(* IEC 61131-3 sources: deprecated-refusr-repo/GP/Main/samples (part 22) *)

(* ---- RND-EXPR_mouse-rusts-agues.st ---- *)
(*
This code implements a randomly grown symbolic expression:

((((!(!(!(xor(xor(IN40 | (xor(xor(IN19, IN3), IN23)), xor(xor(IN26 & IN29, !(IN6)), IN3 & IN48)), xor(xor(IN48 | IN38, !(IN41)), IN9 & IN1)))))) & true) | (xor(xor(!(IN21 & (IN50 | (IN33 & (!(!(IN10)))))), !(IN33)), IN31))) | (!(xor(xor((xor(xor(!(IN26 & (!(!(IN15)))), xor(xor((IN23 | (xor(xor(IN10, IN17), IN38))) | ((IN9 | IN7) | (IN42 & IN18)), (!(IN3)) | (!(IN26 & IN36))), xor(xor(!(IN23), (xor(xor(IN46, IN32), IN13)) | (!(IN45))), IN31))), !(xor(xor(!(xor(xor(IN29, IN29), IN17)), (IN32 | IN36) | (xor(xor(IN34, IN37), true))), xor(xor(IN48 & IN9, xor(xor(IN43, IN49), IN14)), IN2))))) | (!(((xor(xor(!(IN32), xor(xor(IN27, IN24), IN34)), IN7)) & true) | IN46)), !(IN23)), xor(xor(xor(xor((xor(xor((xor(xor(IN42, IN37), IN30)) | IN36, !(IN36)), IN31)) | (!(IN26 | (IN2 | IN28))), (!(IN14)) & (xor(xor((IN45 & IN11) | (xor(xor(IN8, IN48), IN36)), (!(IN36)) & (IN20 & IN4)), !(IN9 & IN11)))), (IN50 | (!(xor(xor(IN12, IN4), IN6)))) | (IN22 & ((IN46 & IN5) & (!(IN41))))), xor(xor(IN41, !(((IN26 & IN16) | (!(IN32))) | ((xor(xor(IN22, IN34), IN14)) & (xor(xor(IN18, IN31), IN36))))), xor(xor((IN8 | (IN9 & IN25)) & (xor(xor(!(IN41), !(IN45)), IN30 & IN43)), (!(IN18 | IN43)) | ((IN39 | IN36) & IN3)), xor(xor(IN44, (xor(xor(IN5, IN21), IN30)) | (xor(xor(IN43, IN17), IN49))), IN30)))), (!(xor(xor(IN44 & (!(IN21)), IN27), (xor(xor(IN34, IN5), IN26)) | (IN38 & IN23)))) | ((!((IN15 | IN19) | (!(IN41)))) & IN20)))))) & (((!((xor(xor(((IN40 & (!(IN13))) | ((!(IN22)) | IN28)) | (xor(xor((IN20 | IN38) & (!(IN15)), !(!(IN14))), true)), (xor(xor(xor(xor(IN5, IN3), IN26 | IN3), xor(xor(true | IN14, !(IN17)), xor(xor(IN17, IN36), IN47))), (xor(xor(IN3, IN48), IN41)) | (IN2 & IN4))) & IN40), ((!(IN6 & IN11)) & (IN26 & (IN27 | IN31))) | (IN49 & (!(xor(xor(IN27, IN28), IN2)))))) | ((xor(xor(!((IN41 | IN16) | (IN35 & IN24)), IN38), xor(xor(!(IN15 & IN10), (IN7 | IN17) | (IN38 & IN35)), xor(xor(IN41 & IN32, IN3 | IN1), !(IN20))))) & (xor(xor((xor(xor(IN6, IN30 | IN35), xor(xor(IN20, IN9), IN29))) & ((IN14 & IN14) & (IN34 | IN49)), IN15), xor(xor(true, !(IN41 & IN2)), (!(IN13)) | (IN24 | true))))))) | IN32) & (xor(xor(IN26, ((((xor(xor(xor(xor(xor(xor(IN9, IN24), IN27), IN45 | IN12), IN10 | IN19), IN7 | (IN12 & IN13)), (!(IN20)) & (!(IN2)))) | (xor(xor((IN20 | IN22) & (IN42 | false), !(IN43 & IN7)), xor(xor(!(IN49), xor(xor(IN31, IN26), IN38)), xor(xor(IN23, IN1), IN3))))) & (((!(IN4 & IN31)) | IN41) & (((xor(xor(IN34, IN47), IN25)) & (xor(xor(IN13, IN11), IN1))) & IN26))) & (!(xor(xor(xor(xor(IN50 & (IN10 | IN31), xor(xor(IN33, xor(xor(IN36, IN43), IN43)), xor(xor(IN21, IN20), IN23))), IN6), ((!(IN48)) | (IN35 & IN49)) & (xor(xor(xor(xor(IN1, IN38), IN48), !(IN17)), IN8 | IN26))), xor(xor((IN23 | IN47) | (xor(xor(IN19, IN38), IN1)), !(IN48)), xor(xor(false, xor(xor(IN31, IN1), IN6)), !(IN34))))))) & (xor(xor(IN9, xor(xor((!((IN29 & IN46) & (!(IN5)))) | IN47, (!((IN45 & IN35) & (!(IN14)))) & IN1), IN14 | (!(IN38)))), xor(xor((!(!(!(IN40)))) & ((xor(xor(!(IN18), IN7), IN17 & IN6)) | (xor(xor(xor(xor(IN12, IN34), IN21), true | IN23), !(IN1)))), !(IN43)), (((IN6 & IN32) | (!(IN11))) & (!(IN24))) & (!(xor(xor(IN36 | IN16, !(IN7)), !(IN30)))))))), (xor(xor(xor(xor((xor(xor(!(IN40 & IN14), xor(xor(!(IN45), xor(xor(IN10, IN14), IN43)), !(IN16))), xor(xor(IN10 | IN17, xor(xor(true, IN13), IN11)), IN4 & IN1))) | IN23, IN43), xor(xor(IN7, !(xor(xor(!(IN30), IN16 | IN10), IN26 | IN18))), !(!(IN42 | IN8)))), ((!(IN46)) & (xor(xor(IN45, xor(xor(!(IN32), xor(xor(IN41, IN14), IN50)), IN22 & IN33)), IN23 & IN27))) & IN4), IN2)) | (!((xor(xor(xor(xor(IN7, xor(xor(IN40, xor(xor(IN42, IN46), IN3)), !(IN41))), (xor(xor(IN5, IN22), IN18)) & (IN47 & IN38)), IN47), IN50)) | ((xor(xor((IN13 & IN49) | (IN6 & IN16), (IN20 & IN30) | (xor(xor(IN22, IN10), IN39))), IN40)) | false))))))

*)

FUNCTION_BLOCK F_CollectInput
  VAR_IN_OUT
      Data : ARRAY[1..50] OF BOOL;
  END_VAR
  VAR_INPUT
      TICK  : BOOL := 0;
      IN1   : BOOL := 0;
      IN2   : BOOL := 0;
      IN3   : BOOL := 0;
      IN4   : BOOL := 0;
      IN5   : BOOL := 0;
      RESET : BOOL := FALSE;
  END_VAR
  VAR_OUTPUT
      Finished : BOOL;
  END_VAR
  VAR
      j    : USINT := 1;
      tock : BOOL  := 0;
  END_VAR
  IF NOT RESET AND tock = NOT TICK THEN
      Data[j]   := IN1;
      Data[j+1] := IN2;
      Data[j+2] := IN3;
      Data[j+3] := IN4;
      Data[j+4] := IN5;
      j := j + 5;
      tock := TICK;
  ELSE
      j := 1;
      tock := 0;
  END_IF;
  Finished := (j > 50);
END_FUNCTION_BLOCK

PROGRAM Boiler
  VAR
    Data  : ARRAY[1..50] OF BOOL;
    Ready : BOOL;
    CollectInput : F_CollectInput;
  END_VAR
  VAR
    TICK     AT %IX1.0 : BOOL;
    IN1      AT %IX0.3 : BOOL;
    IN2      AT %IX0.4 : BOOL;
    IN3      AT %IX0.5 : BOOL;
    IN4      AT %IX0.6 : BOOL;
    IN5      AT %IX0.7 : BOOL;
    OutReady AT %QX0.0 : BOOL := FALSE;
    FeedNext AT %QX0.1 : BOOL := FALSE;
    Out      AT %QX0.2 : BOOL;
  END_VAR
  CollectInput(TICK:=TICK, IN1:=IN1, IN2:=IN2, IN3:=IN3, IN4:=IN4, IN5:=IN5);
  Ready := CollectInput.Finished;
  FeedNext := 1;
  IF Ready THEN
    Out := (((((NOT (NOT (NOT (((Data[40] OR ((Data[19] XOR Data[3]) XOR Data[23])) XOR (((Data[26] AND Data[29]) XOR (NOT Data[6])) XOR (Data[3] AND Data[48]))) XOR (((Data[48] OR Data[38]) XOR (NOT Data[41])) XOR (Data[9] AND Data[1])))))) AND TRUE) OR (((NOT (Data[21] AND (Data[50] OR (Data[33] AND (NOT (NOT Data[10])))))) XOR (NOT Data[33])) XOR Data[31])) OR (NOT ((((((NOT (Data[26] AND (NOT (NOT Data[15])))) XOR ((((Data[23] OR ((Data[10] XOR Data[17]) XOR Data[38])) OR ((Data[9] OR Data[7]) OR (Data[42] AND Data[18]))) XOR ((NOT Data[3]) OR (NOT (Data[26] AND Data[36])))) XOR (((NOT Data[23]) XOR (((Data[46] XOR Data[32]) XOR Data[13]) OR (NOT Data[45]))) XOR Data[31]))) XOR (NOT (((NOT ((Data[29] XOR Data[29]) XOR Data[17])) XOR ((Data[32] OR Data[36]) OR ((Data[34] XOR Data[37]) XOR TRUE))) XOR (((Data[48] AND Data[9]) XOR ((Data[43] XOR Data[49]) XOR Data[14])) XOR Data[2])))) OR (NOT (((((NOT Data[32]) XOR ((Data[27] XOR Data[24]) XOR Data[34])) XOR Data[7]) AND TRUE) OR Data[46]))) XOR (NOT Data[23])) XOR ((((((((((Data[42] XOR Data[37]) XOR Data[30]) OR Data[36]) XOR (NOT Data[36])) XOR Data[31]) OR (NOT (Data[26] OR (Data[2] OR Data[28])))) XOR ((NOT Data[14]) AND ((((Data[45] AND Data[11]) OR ((Data[8] XOR Data[48]) XOR Data[36])) XOR ((NOT Data[36]) AND (Data[20] AND Data[4]))) XOR (NOT (Data[9] AND Data[11]))))) XOR ((Data[50] OR (NOT ((Data[12] XOR Data[4]) XOR Data[6]))) OR (Data[22] AND ((Data[46] AND Data[5]) AND (NOT Data[41]))))) XOR ((Data[41] XOR (NOT (((Data[26] AND Data[16]) OR (NOT Data[32])) OR (((Data[22] XOR Data[34]) XOR Data[14]) AND ((Data[18] XOR Data[31]) XOR Data[36]))))) XOR ((((Data[8] OR (Data[9] AND Data[25])) AND (((NOT Data[41]) XOR (NOT Data[45])) XOR (Data[30] AND Data[43]))) XOR ((NOT (Data[18] OR Data[43])) OR ((Data[39] OR Data[36]) AND Data[3]))) XOR ((Data[44] XOR (((Data[5] XOR Data[21]) XOR Data[30]) OR ((Data[43] XOR Data[17]) XOR Data[49]))) XOR Data[30])))) XOR ((NOT (((Data[44] AND (NOT Data[21])) XOR Data[27]) XOR (((Data[34] XOR Data[5]) XOR Data[26]) OR (Data[38] AND Data[23])))) OR ((NOT ((Data[15] OR Data[19]) OR (NOT Data[41]))) AND Data[20])))))) AND (((NOT ((((((Data[40] AND (NOT Data[13])) OR ((NOT Data[22]) OR Data[28])) OR ((((Data[20] OR Data[38]) AND (NOT Data[15])) XOR (NOT (NOT Data[14]))) XOR TRUE)) XOR (((((Data[5] XOR Data[3]) XOR (Data[26] OR Data[3])) XOR (((TRUE OR Data[14]) XOR (NOT Data[17])) XOR ((Data[17] XOR Data[36]) XOR Data[47]))) XOR (((Data[3] XOR Data[48]) XOR Data[41]) OR (Data[2] AND Data[4]))) AND Data[40])) XOR (((NOT (Data[6] AND Data[11])) AND (Data[26] AND (Data[27] OR Data[31]))) OR (Data[49] AND (NOT ((Data[27] XOR Data[28]) XOR Data[2]))))) OR ((((NOT ((Data[41] OR Data[16]) OR (Data[35] AND Data[24]))) XOR Data[38]) XOR (((NOT (Data[15] AND Data[10])) XOR ((Data[7] OR Data[17]) OR (Data[38] AND Data[35]))) XOR (((Data[41] AND Data[32]) XOR (Data[3] OR Data[1])) XOR (NOT Data[20])))) AND (((((Data[6] XOR (Data[30] OR Data[35])) XOR ((Data[20] XOR Data[9]) XOR Data[29])) AND ((Data[14] AND Data[14]) AND (Data[34] OR Data[49]))) XOR Data[15]) XOR ((TRUE XOR (NOT (Data[41] AND Data[2]))) XOR ((NOT Data[13]) OR (Data[24] OR TRUE))))))) OR Data[32]) AND ((Data[26] XOR ((((((((((Data[9] XOR Data[24]) XOR Data[27]) XOR (Data[45] OR Data[12])) XOR (Data[10] OR Data[19])) XOR (Data[7] OR (Data[12] AND Data[13]))) XOR ((NOT Data[20]) AND (NOT Data[2]))) OR ((((Data[20] OR Data[22]) AND (Data[42] OR FALSE)) XOR (NOT (Data[43] AND Data[7]))) XOR (((NOT Data[49]) XOR ((Data[31] XOR Data[26]) XOR Data[38])) XOR ((Data[23] XOR Data[1]) XOR Data[3])))) AND (((NOT (Data[4] AND Data[31])) OR Data[41]) AND ((((Data[34] XOR Data[47]) XOR Data[25]) AND ((Data[13] XOR Data[11]) XOR Data[1])) AND Data[26]))) AND (NOT (((((Data[50] AND (Data[10] OR Data[31])) XOR ((Data[33] XOR ((Data[36] XOR Data[43]) XOR Data[43])) XOR ((Data[21] XOR Data[20]) XOR Data[23]))) XOR Data[6]) XOR (((NOT Data[48]) OR (Data[35] AND Data[49])) AND ((((Data[1] XOR Data[38]) XOR Data[48]) XOR (NOT Data[17])) XOR (Data[8] OR Data[26])))) XOR ((((Data[23] OR Data[47]) OR ((Data[19] XOR Data[38]) XOR Data[1])) XOR (NOT Data[48])) XOR ((FALSE XOR ((Data[31] XOR Data[1]) XOR Data[6])) XOR (NOT Data[34])))))) AND ((Data[9] XOR ((((NOT ((Data[29] AND Data[46]) AND (NOT Data[5]))) OR Data[47]) XOR ((NOT ((Data[45] AND Data[35]) AND (NOT Data[14]))) AND Data[1])) XOR (Data[14] OR (NOT Data[38])))) XOR ((((NOT (NOT (NOT Data[40]))) AND ((((NOT Data[18]) XOR Data[7]) XOR (Data[17] AND Data[6])) OR ((((Data[12] XOR Data[34]) XOR Data[21]) XOR (TRUE OR Data[23])) XOR (NOT Data[1])))) XOR (NOT Data[43])) XOR ((((Data[6] AND Data[32]) OR (NOT Data[11])) AND (NOT Data[24])) AND (NOT (((Data[36] OR Data[16]) XOR (NOT Data[7])) XOR (NOT Data[30])))))))) XOR (((((((((NOT (Data[40] AND Data[14])) XOR (((NOT Data[45]) XOR ((Data[10] XOR Data[14]) XOR Data[43])) XOR (NOT Data[16]))) XOR (((Data[10] OR Data[17]) XOR ((TRUE XOR Data[13]) XOR Data[11])) XOR (Data[4] AND Data[1]))) OR Data[23]) XOR Data[43]) XOR ((Data[7] XOR (NOT (((NOT Data[30]) XOR (Data[16] OR Data[10])) XOR (Data[26] OR Data[18])))) XOR (NOT (NOT (Data[42] OR Data[8]))))) XOR (((NOT Data[46]) AND ((Data[45] XOR (((NOT Data[32]) XOR ((Data[41] XOR Data[14]) XOR Data[50])) XOR (Data[22] AND Data[33]))) XOR (Data[23] AND Data[27]))) AND Data[4])) XOR Data[2]) OR (NOT (((((Data[7] XOR ((Data[40] XOR ((Data[42] XOR Data[46]) XOR Data[3])) XOR (NOT Data[41]))) XOR (((Data[5] XOR Data[22]) XOR Data[18]) AND (Data[47] AND Data[38]))) XOR Data[47]) XOR Data[50]) OR (((((Data[13] AND Data[49]) OR (Data[6] AND Data[16])) XOR ((Data[20] AND Data[30]) OR ((Data[22] XOR Data[10]) XOR Data[39]))) XOR Data[40]) OR FALSE)))))));
    OutReady := 1;
    CollectInput(RESET:=TRUE);
  END_IF;
END_PROGRAM

CONFIGURATION Config0
  RESOURCE Res0 ON PLC
    TASK task0(INTERVAL := T#20ms,PRIORITY := 0);
    PROGRAM instance0 WITH task0 : Boiler;
  END_RESOURCE
END_CONFIGURATION

(* ---- RND-EXPR_musky-murky-tasty.st ---- *)
(*
This code implements a randomly grown symbolic expression:

xor(xor(IN21, xor(xor(!(xor(xor(!(((IN33 | (!(xor(xor(IN43, IN17), IN41)))) | (((IN24 & IN36) | IN2) & ((IN39 & IN3) & (!(IN44))))) | (!(!(xor(xor(IN35 & IN26, IN42 & IN24), !(IN4)))))), (xor(xor(((!(IN11 & IN23)) & (!(IN3 | true))) | IN47, xor(xor(xor(xor(xor(xor(!(IN14), !(IN37)), xor(xor(IN10, IN8), IN22)), xor(xor(xor(xor(IN29, IN50), IN7), !(IN35)), IN3 & IN45)), IN46 | (IN26 | IN44)), IN38), !((IN41 | IN26) | (IN19 | IN47)))), !(((!(IN41)) & IN13) & (xor(xor(IN49 | IN49, xor(xor(IN43, IN4), IN24)), !(IN49)))))) | IN18), (((IN32 & ((!(IN18)) | (xor(xor(IN33, IN30), IN29)))) & (xor(xor(IN7, (IN4 | IN26) | (IN25 & IN38)), (IN25 & IN24) & (xor(xor(IN27, false), IN39))))) | (xor(xor(((xor(xor(IN7, IN42), IN10)) | IN32) & (xor(xor(IN17, xor(xor(IN39, IN31), IN37)), IN7)), !(xor(xor(!(IN43), !(IN16)), IN50 | IN35))), (xor(xor(IN19, IN4 | IN18), IN36)) & ((!(IN22)) | IN19)))) | IN21)), IN44), xor(xor(((xor(xor(!(xor(xor(!(IN35 | IN45), (!(IN27)) & (IN43 & IN44)), xor(xor(IN46, IN15 & IN22), !(IN33)))), !(!((!(IN36)) | (IN16 | IN14)))), IN23 | (xor(xor(IN10 & IN4, xor(xor(xor(xor(IN34, IN37), IN13), IN47), !(IN31))), xor(xor(IN12 & IN11, IN12 | IN18), !(IN39)))))) | (!(!(!(xor(xor(xor(xor(IN14, IN14), IN19), IN45 & IN38), IN15)))))) | ((xor(xor((((IN33 | IN36) | (!(IN20))) & (IN33 & (IN33 & IN33))) | (xor(xor(IN45 | (IN8 & IN21), xor(xor(xor(xor(IN31, IN46), IN43), xor(xor(IN48, IN2), IN12)), IN28)), !(IN49))), xor(xor(xor(xor(xor(xor(!(IN27), xor(xor(IN16, IN38), IN22)), IN26 | IN35), !(IN3 & IN47)), !(IN42 | IN28)), !(IN31)), !(IN39))), (xor(xor((xor(xor(IN27, IN35), IN17)) & (IN13 & IN30), IN15), !(xor(xor(IN39, IN29), IN46)))) | (((!(IN47)) | (IN22 | IN32)) | (!(IN29 | IN7))))) & IN13), IN3 & (!(xor(xor(xor(xor((!(!(IN22))) & (!(IN22 | IN20)), ((IN13 & IN28) & (!(IN27))) | (xor(xor(!(IN27), !(IN36)), IN20 | IN44))), IN19), ((xor(xor(xor(xor(IN7, IN21), IN13), IN40 | IN47), !(IN32))) | (xor(xor(IN29 | IN15, !(IN26)), !(IN27)))) | ((xor(xor(IN27 | IN24, xor(xor(IN27, IN23), IN6)), !(IN47))) & ((IN12 | IN31) | (!(IN16))))), (!(!(IN46))) & IN15)))), !(xor(xor(xor(xor((!(!(!(IN11)))) & ((!(false | IN24)) & (xor(xor(!(IN48), xor(xor(IN41, true), IN47)), !(IN11)))), IN36), (IN35 & (xor(xor(xor(xor(IN40, IN32), IN38), xor(xor(IN44, IN29), IN18)), false | IN50))) | (((IN36 & IN23) | (!(IN9))) & (!(IN39 | IN43)))), !(((!(xor(xor(IN29, IN9), IN19))) & ((IN6 & IN41) | (IN20 & IN14))) | (!(true & (IN40 | IN30))))), !(((!(IN16)) & (xor(xor(xor(xor(IN46, IN30), IN2), !(IN40)), false))) | (xor(xor(!(IN20 | IN25), !(IN50 | IN1)), IN42)))))))), IN7)

*)

FUNCTION_BLOCK F_CollectInput
  VAR_IN_OUT
      Data : ARRAY[1..50] OF BOOL;
  END_VAR
  VAR_INPUT
      TICK  : BOOL := 0;
      IN1   : BOOL := 0;
      IN2   : BOOL := 0;
      IN3   : BOOL := 0;
      IN4   : BOOL := 0;
      IN5   : BOOL := 0;
      RESET : BOOL := FALSE;
  END_VAR
  VAR_OUTPUT
      Finished : BOOL;
  END_VAR
  VAR
      j    : USINT := 1;
      tock : BOOL  := 0;
  END_VAR
  IF NOT RESET AND tock = NOT TICK THEN
      Data[j]   := IN1;
      Data[j+1] := IN2;
      Data[j+2] := IN3;
      Data[j+3] := IN4;
      Data[j+4] := IN5;
      j := j + 5;
      tock := TICK;
  ELSE
      j := 1;
      tock := 0;
  END_IF;
  Finished := (j > 50);
END_FUNCTION_BLOCK

PROGRAM Boiler
  VAR
    Data  : ARRAY[1..50] OF BOOL;
    Ready : BOOL;
    CollectInput : F_CollectInput;
  END_VAR
  VAR
    TICK     AT %IX1.0 : BOOL;
    IN1      AT %IX0.3 : BOOL;
    IN2      AT %IX0.4 : BOOL;
    IN3      AT %IX0.5 : BOOL;
    IN4      AT %IX0.6 : BOOL;
    IN5      AT %IX0.7 : BOOL;
    OutReady AT %QX0.0 : BOOL := FALSE;
    FeedNext AT %QX0.1 : BOOL := FALSE;
    Out      AT %QX0.2 : BOOL;
  END_VAR
  CollectInput(TICK:=TICK, IN1:=IN1, IN2:=IN2, IN3:=IN3, IN4:=IN4, IN5:=IN5);
  Ready := CollectInput.Finished;
  FeedNext := 1;
  IF Ready THEN
    Out := ((Data[21] XOR (((NOT (((NOT (((Data[33] OR (NOT ((Data[43] XOR Data[17]) XOR Data[41]))) OR (((Data[24] AND Data[36]) OR Data[2]) AND ((Data[39] AND Data[3]) AND (NOT Data[44])))) OR (NOT (NOT (((Data[35] AND Data[26]) XOR (Data[42] AND Data[24])) XOR (NOT Data[4])))))) XOR ((((((NOT (Data[11] AND Data[23])) AND (NOT (Data[3] OR TRUE))) OR Data[47]) XOR (((((((NOT Data[14]) XOR (NOT Data[37])) XOR ((Data[10] XOR Data[8]) XOR Data[22])) XOR ((((Data[29] XOR Data[50]) XOR Data[7]) XOR (NOT Data[35])) XOR (Data[3] AND Data[45]))) XOR (Data[46] OR (Data[26] OR Data[44]))) XOR Data[38]) XOR (NOT ((Data[41] OR Data[26]) OR (Data[19] OR Data[47]))))) XOR (NOT (((NOT Data[41]) AND Data[13]) AND (((Data[49] OR Data[49]) XOR ((Data[43] XOR Data[4]) XOR Data[24])) XOR (NOT Data[49]))))) OR Data[18])) XOR ((((Data[32] AND ((NOT Data[18]) OR ((Data[33] XOR Data[30]) XOR Data[29]))) AND ((Data[7] XOR ((Data[4] OR Data[26]) OR (Data[25] AND Data[38]))) XOR ((Data[25] AND Data[24]) AND ((Data[27] XOR FALSE) XOR Data[39])))) OR ((((((Data[7] XOR Data[42]) XOR Data[10]) OR Data[32]) AND ((Data[17] XOR ((Data[39] XOR Data[31]) XOR Data[37])) XOR Data[7])) XOR (NOT (((NOT Data[43]) XOR (NOT Data[16])) XOR (Data[50] OR Data[35])))) XOR (((Data[19] XOR (Data[4] OR Data[18])) XOR Data[36]) AND ((NOT Data[22]) OR Data[19])))) OR Data[21]))) XOR Data[44]) XOR (((((((NOT (((NOT (Data[35] OR Data[45])) XOR ((NOT Data[27]) AND (Data[43] AND Data[44]))) XOR ((Data[46] XOR (Data[15] AND Data[22])) XOR (NOT Data[33])))) XOR (NOT (NOT ((NOT Data[36]) OR (Data[16] OR Data[14]))))) XOR (Data[23] OR (((Data[10] AND Data[4]) XOR ((((Data[34] XOR Data[37]) XOR Data[13]) XOR Data[47]) XOR (NOT Data[31]))) XOR (((Data[12] AND Data[11]) XOR (Data[12] OR Data[18])) XOR (NOT Data[39]))))) OR (NOT (NOT (NOT ((((Data[14] XOR Data[14]) XOR Data[19]) XOR (Data[45] AND Data[38])) XOR Data[15]))))) OR (((((((Data[33] OR Data[36]) OR (NOT Data[20])) AND (Data[33] AND (Data[33] AND Data[33]))) OR (((Data[45] OR (Data[8] AND Data[21])) XOR ((((Data[31] XOR Data[46]) XOR Data[43]) XOR ((Data[48] XOR Data[2]) XOR Data[12])) XOR Data[28])) XOR (NOT Data[49]))) XOR (((((((NOT Data[27]) XOR ((Data[16] XOR Data[38]) XOR Data[22])) XOR (Data[26] OR Data[35])) XOR (NOT (Data[3] AND Data[47]))) XOR (NOT (Data[42] OR Data[28]))) XOR (NOT Data[31])) XOR (NOT Data[39]))) XOR ((((((Data[27] XOR Data[35]) XOR Data[17]) AND (Data[13] AND Data[30])) XOR Data[15]) XOR (NOT ((Data[39] XOR Data[29]) XOR Data[46]))) OR (((NOT Data[47]) OR (Data[22] OR Data[32])) OR (NOT (Data[29] OR Data[7]))))) AND Data[13])) XOR (Data[3] AND (NOT ((((((NOT (NOT Data[22])) AND (NOT (Data[22] OR Data[20]))) XOR (((Data[13] AND Data[28]) AND (NOT Data[27])) OR (((NOT Data[27]) XOR (NOT Data[36])) XOR (Data[20] OR Data[44])))) XOR Data[19]) XOR ((((((Data[7] XOR Data[21]) XOR Data[13]) XOR (Data[40] OR Data[47])) XOR (NOT Data[32])) OR (((Data[29] OR Data[15]) XOR (NOT Data[26])) XOR (NOT Data[27]))) OR ((((Data[27] OR Data[24]) XOR ((Data[27] XOR Data[23]) XOR Data[6])) XOR (NOT Data[47])) AND ((Data[12] OR Data[31]) OR (NOT Data[16]))))) XOR ((NOT (NOT Data[46])) AND Data[15]))))) XOR (NOT ((((((NOT (NOT (NOT Data[11]))) AND ((NOT (FALSE OR Data[24])) AND (((NOT Data[48]) XOR ((Data[41] XOR TRUE) XOR Data[47])) XOR (NOT Data[11])))) XOR Data[36]) XOR ((Data[35] AND ((((Data[40] XOR Data[32]) XOR Data[38]) XOR ((Data[44] XOR Data[29]) XOR Data[18])) XOR (FALSE OR Data[50]))) OR (((Data[36] AND Data[23]) OR (NOT Data[9])) AND (NOT (Data[39] OR Data[43]))))) XOR (NOT (((NOT ((Data[29] XOR Data[9]) XOR Data[19])) AND ((Data[6] AND Data[41]) OR (Data[20] AND Data[14]))) OR (NOT (TRUE AND (Data[40] OR Data[30])))))) XOR (NOT (((NOT Data[16]) AND ((((Data[46] XOR Data[30]) XOR Data[2]) XOR (NOT Data[40])) XOR FALSE)) OR (((NOT (Data[20] OR Data[25])) XOR (NOT (Data[50] OR Data[1]))) XOR Data[42])))))))) XOR Data[7]);
    OutReady := 1;
    CollectInput(RESET:=TRUE);
  END_IF;
END_PROGRAM

CONFIGURATION Config0
  RESOURCE Res0 ON PLC
    TASK task0(INTERVAL := T#20ms,PRIORITY := 0);
    PROGRAM instance0 WITH task0 : Boiler;
  END_RESOURCE
END_CONFIGURATION

(* ---- RND-EXPR_organ-ionic-vodka.st ---- *)
(*
This code implements a randomly grown symbolic expression:

(!(!((!((xor(xor((!(IN50 & IN40)) | ((xor(xor(IN25, IN48), IN45)) | (!(IN5))), (xor(xor(!(IN44), IN40 | IN25), !(IN39))) | ((xor(xor(IN39, IN46), IN37)) | (IN1 | IN32))), !(xor(xor(xor(xor(IN6, IN50), IN24), xor(xor(IN17, true), IN37)), xor(xor(true, IN48), IN13))))) & ((IN35 & (!(IN47))) & ((xor(xor(IN23 & IN22, IN2 & IN37), IN6 | true)) | (xor(xor(IN40, IN45 | IN9), IN42 & IN5)))))) | (xor(xor((((xor(xor(xor(xor(IN25, IN3), IN34), xor(xor(IN46, IN17), IN18)), IN23 & IN14)) | ((!(IN46)) & (IN8 | IN2))) & (!((xor(xor(IN25, IN19), IN42)) & (!(IN16))))) & ((xor(xor(xor(xor(true & IN31, !(IN14)), IN7 & IN30), IN21), IN18)) & ((!(IN16 & IN29)) | (!(!(IN28))))), ((xor(xor(xor(xor(IN37 | IN10, !(IN13)), IN30 | true), (xor(xor(IN25, IN7), IN15)) | (IN1 & IN31)), (xor(xor(IN7, IN29), IN14)) | (IN38 & IN27))) & (!((IN20 & IN25) & (xor(xor(IN18, IN13), IN34))))) | IN29), IN38))))) & ((xor(xor(xor(xor(IN2 | (IN37 | (!(xor(xor(IN47, IN31), xor(xor(xor(xor(IN29, IN18), IN30), IN33 | IN32), IN21 | IN40))))), !((!((!(IN43)) & (xor(xor(IN15, IN37), IN16 & IN49)))) & (xor(xor((!(!(IN16))) | (!(IN31 & IN33)), !((IN43 & IN11) & (IN30 | IN6))), !(xor(xor(!(IN9), IN21 & IN34), xor(xor(IN7, true), IN4))))))), ((IN22 | IN45) | (!((xor(xor(IN18, !(IN9)), !(IN13))) & (xor(xor(IN25, !(IN31)), IN20))))) & (xor(xor((((IN37 & IN22) | (IN9 | IN25)) & IN48) & (((IN20 & IN20) & (IN13 | IN8)) & (IN11 & IN7)), (IN3 | ((!(IN40)) & (!(IN33)))) | ((xor(xor(IN15, xor(xor(false, IN49), IN27)), xor(xor(IN36, IN19), IN36))) & (xor(xor(IN24, IN43 & IN35), IN8 & IN10)))), ((xor(xor(false, xor(xor(IN43, IN33), IN12)), IN45 | IN19)) & (xor(xor(IN35 & IN39, !(IN29)), IN4))) & (xor(xor(IN21, (!(IN34)) & (xor(xor(IN7, IN20), IN8))), (IN27 & IN41) & (IN2 | IN24)))))), !(IN41)), xor(xor(false, ((!(IN50 & IN2)) & (IN15 | (((IN18 & IN46) & (false & IN39)) & ((IN36 | IN28) | (!(IN19)))))) | (xor(xor(false & (((IN23 | IN12) | (IN9 & IN49)) & (!(IN26 | IN44))), IN48), IN21 | ((xor(xor(IN35, IN6 | false), IN9 & IN13)) | ((!(IN20)) & (!(IN23))))))), !(!(!(((IN21 & IN20) | (xor(xor(IN35, IN5), IN47))) & (xor(xor(IN4 | IN35, xor(xor(IN40, IN19), IN43)), IN44)))))))) & (!((xor(xor(IN39, IN23), IN3)) | ((xor(xor(IN25, !(IN42)), IN31)) | (xor(xor(((!(IN43 & IN30)) & (IN12 & IN48)) & ((!(IN44)) | IN42), (xor(xor(xor(xor(IN38, IN24 | IN20), IN1), xor(xor(true, IN36 | IN9), IN40 & IN33)), (IN44 & IN41) | (IN44 | IN48))) & true), IN17))))))

*)

FUNCTION_BLOCK F_CollectInput
  VAR_IN_OUT
      Data : ARRAY[1..50] OF BOOL;
  END_VAR
  VAR_INPUT
      TICK  : BOOL := 0;
      IN1   : BOOL := 0;
      IN2   : BOOL := 0;
      IN3   : BOOL := 0;
      IN4   : BOOL := 0;
      IN5   : BOOL := 0;
      RESET : BOOL := FALSE;
  END_VAR
  VAR_OUTPUT
      Finished : BOOL;
  END_VAR
  VAR
      j    : USINT := 1;
      tock : BOOL  := 0;
  END_VAR
  IF NOT RESET AND tock = NOT TICK THEN
      Data[j]   := IN1;
      Data[j+1] := IN2;
      Data[j+2] := IN3;
      Data[j+3] := IN4;
      Data[j+4] := IN5;
      j := j + 5;
      tock := TICK;
  ELSE
      j := 1;
      tock := 0;
  END_IF;
  Finished := (j > 50);
END_FUNCTION_BLOCK

PROGRAM Boiler
  VAR
    Data  : ARRAY[1..50] OF BOOL;
    Ready : BOOL;
    CollectInput : F_CollectInput;
  END_VAR
  VAR
    TICK     AT %IX1.0 : BOOL;
    IN1      AT %IX0.3 : BOOL;
    IN2      AT %IX0.4 : BOOL;
    IN3      AT %IX0.5 : BOOL;
    IN4      AT %IX0.6 : BOOL;
    IN5      AT %IX0.7 : BOOL;
    OutReady AT %QX0.0 : BOOL := FALSE;
    FeedNext AT %QX0.1 : BOOL := FALSE;
    Out      AT %QX0.2 : BOOL;
  END_VAR
  CollectInput(TICK:=TICK, IN1:=IN1, IN2:=IN2, IN3:=IN3, IN4:=IN4, IN5:=IN5);
  Ready := CollectInput.Finished;
  FeedNext := 1;
  IF Ready THEN
    Out := ((NOT (NOT ((NOT (((((NOT (Data[50] AND Data[40])) OR (((Data[25] XOR Data[48]) XOR Data[45]) OR (NOT Data[5]))) XOR ((((NOT Data[44]) XOR (Data[40] OR Data[25])) XOR (NOT Data[39])) OR (((Data[39] XOR Data[46]) XOR Data[37]) OR (Data[1] OR Data[32])))) XOR (NOT ((((Data[6] XOR Data[50]) XOR Data[24]) XOR ((Data[17] XOR TRUE) XOR Data[37])) XOR ((TRUE XOR Data[48]) XOR Data[13])))) AND ((Data[35] AND (NOT Data[47])) AND ((((Data[23] AND Data[22]) XOR (Data[2] AND Data[37])) XOR (Data[6] OR TRUE)) OR ((Data[40] XOR (Data[45] OR Data[9])) XOR (Data[42] AND Data[5])))))) OR (((((((((Data[25] XOR Data[3]) XOR Data[34]) XOR ((Data[46] XOR Data[17]) XOR Data[18])) XOR (Data[23] AND Data[14])) OR ((NOT Data[46]) AND (Data[8] OR Data[2]))) AND (NOT (((Data[25] XOR Data[19]) XOR Data[42]) AND (NOT Data[16])))) AND ((((((TRUE AND Data[31]) XOR (NOT Data[14])) XOR (Data[7] AND Data[30])) XOR Data[21]) XOR Data[18]) AND ((NOT (Data[16] AND Data[29])) OR (NOT (NOT Data[28]))))) XOR (((((((Data[37] OR Data[10]) XOR (NOT Data[13])) XOR (Data[30] OR TRUE)) XOR (((Data[25] XOR Data[7]) XOR Data[15]) OR (Data[1] AND Data[31]))) XOR (((Data[7] XOR Data[29]) XOR Data[14]) OR (Data[38] AND Data[27]))) AND (NOT ((Data[20] AND Data[25]) AND ((Data[18] XOR Data[13]) XOR Data[34])))) OR Data[29])) XOR Data[38])))) AND ((((((Data[2] OR (Data[37] OR (NOT ((Data[47] XOR Data[31]) XOR ((((Data[29] XOR Data[18]) XOR Data[30]) XOR (Data[33] OR Data[32])) XOR (Data[21] OR Data[40])))))) XOR (NOT ((NOT ((NOT Data[43]) AND ((Data[15] XOR Data[37]) XOR (Data[16] AND Data[49])))) AND ((((NOT (NOT Data[16])) OR (NOT (Data[31] AND Data[33]))) XOR (NOT ((Data[43] AND Data[11]) AND (Data[30] OR Data[6])))) XOR (NOT (((NOT Data[9]) XOR (Data[21] AND Data[34])) XOR ((Data[7] XOR TRUE) XOR Data[4]))))))) XOR (((Data[22] OR Data[45]) OR (NOT (((Data[18] XOR (NOT Data[9])) XOR (NOT Data[13])) AND ((Data[25] XOR (NOT Data[31])) XOR Data[20])))) AND ((((((Data[37] AND Data[22]) OR (Data[9] OR Data[25])) AND Data[48]) AND (((Data[20] AND Data[20]) AND (Data[13] OR Data[8])) AND (Data[11] AND Data[7]))) XOR ((Data[3] OR ((NOT Data[40]) AND (NOT Data[33]))) OR (((Data[15] XOR ((FALSE XOR Data[49]) XOR Data[27])) XOR ((Data[36] XOR Data[19]) XOR Data[36])) AND ((Data[24] XOR (Data[43] AND Data[35])) XOR (Data[8] AND Data[10]))))) XOR ((((FALSE XOR ((Data[43] XOR Data[33]) XOR Data[12])) XOR (Data[45] OR Data[19])) AND (((Data[35] AND Data[39]) XOR (NOT Data[29])) XOR Data[4])) AND ((Data[21] XOR ((NOT Data[34]) AND ((Data[7] XOR Data[20]) XOR Data[8]))) XOR ((Data[27] AND Data[41]) AND (Data[2] OR Data[24]))))))) XOR (NOT Data[41])) XOR ((FALSE XOR (((NOT (Data[50] AND Data[2])) AND (Data[15] OR (((Data[18] AND Data[46]) AND (FALSE AND Data[39])) AND ((Data[36] OR Data[28]) OR (NOT Data[19]))))) OR (((FALSE AND (((Data[23] OR Data[12]) OR (Data[9] AND Data[49])) AND (NOT (Data[26] OR Data[44])))) XOR Data[48]) XOR (Data[21] OR (((Data[35] XOR (Data[6] OR FALSE)) XOR (Data[9] AND Data[13])) OR ((NOT Data[20]) AND (NOT Data[23]))))))) XOR (NOT (NOT (NOT (((Data[21] AND Data[20]) OR ((Data[35] XOR Data[5]) XOR Data[47])) AND (((Data[4] OR Data[35]) XOR ((Data[40] XOR Data[19]) XOR Data[43])) XOR Data[44]))))))) AND (NOT (((Data[39] XOR Data[23]) XOR Data[3]) OR (((Data[25] XOR (NOT Data[42])) XOR Data[31]) OR (((((NOT (Data[43] AND Data[30])) AND (Data[12] AND Data[48])) AND ((NOT Data[44]) OR Data[42])) XOR (((((Data[38] XOR (Data[24] OR Data[20])) XOR Data[1]) XOR ((TRUE XOR (Data[36] OR Data[9])) XOR (Data[40] AND Data[33]))) XOR ((Data[44] AND Data[41]) OR (Data[44] OR Data[48]))) AND TRUE)) XOR Data[17]))))));
    OutReady := 1;
    CollectInput(RESET:=TRUE);
  END_IF;
END_PROGRAM

CONFIGURATION Config0
  RESOURCE Res0 ON PLC
    TASK task0(INTERVAL := T#20ms,PRIORITY := 0);
    PROGRAM instance0 WITH task0 : Boiler;
  END_RESOURCE
END_CONFIGURATION

(* ---- RND-EXPR_parch-pouch-email.st ---- *)
(*
This code implements a randomly grown symbolic expression:

(((((false & ((((IN32 | IN11) | (IN6 | IN33)) | (IN37 | (!(IN33)))) | (((IN45 | IN22) | (!(IN44))) | (!(IN47))))) | (!(!(IN28)))) & (xor(xor(IN24, xor(xor(IN3 & (xor(xor((IN19 & IN6) & (xor(xor(IN45, IN48), IN8)), xor(xor(!(IN33), IN26 & IN41), IN48)), xor(xor(xor(xor(IN48, IN4), IN30), IN38 & IN7), IN2 & IN27))), (((!(IN46)) & (IN25 & IN22)) | IN3) & IN14), ((!(xor(xor(IN32, IN14), IN46))) | IN41) & ((!(IN32 | IN6)) & (!(!(IN48)))))), !((((xor(xor(IN18, IN35), IN47)) | IN25) | (xor(xor(IN1 | IN9, IN12 & false), true))) & (xor(xor(IN26 | (IN11 & IN20), IN14), !(IN41))))))) | IN15) | (!(!(IN18)))) | IN14

*)

FUNCTION_BLOCK F_CollectInput
  VAR_IN_OUT
      Data : ARRAY[1..50] OF BOOL;
  END_VAR
  VAR_INPUT
      TICK  : BOOL := 0;
      IN1   : BOOL := 0;
      IN2   : BOOL := 0;
      IN3   : BOOL := 0;
      IN4   : BOOL := 0;
      IN5   : BOOL := 0;
      RESET : BOOL := FALSE;
  END_VAR
  VAR_OUTPUT
      Finished : BOOL;
  END_VAR
  VAR
      j    : USINT := 1;
      tock : BOOL  := 0;
  END_VAR
  IF NOT RESET AND tock = NOT TICK THEN
      Data[j]   := IN1;
      Data[j+1] := IN2;
      Data[j+2] := IN3;
      Data[j+3] := IN4;
      Data[j+4] := IN5;
      j := j + 5;
      tock := TICK;
  ELSE
      j := 1;
      tock := 0;
  END_IF;
  Finished := (j > 50);
END_FUNCTION_BLOCK

PROGRAM Boiler
  VAR
    Data  : ARRAY[1..50] OF BOOL;
    Ready : BOOL;
    CollectInput : F_CollectInput;
  END_VAR
  VAR
    TICK     AT %IX1.0 : BOOL;
    IN1      AT %IX0.3 : BOOL;
    IN2      AT %IX0.4 : BOOL;
    IN3      AT %IX0.5 : BOOL;
    IN4      AT %IX0.6 : BOOL;
    IN5      AT %IX0.7 : BOOL;
    OutReady AT %QX0.0 : BOOL := FALSE;
    FeedNext AT %QX0.1 : BOOL := FALSE;
    Out      AT %QX0.2 : BOOL;
  END_VAR
  CollectInput(TICK:=TICK, IN1:=IN1, IN2:=IN2, IN3:=IN3, IN4:=IN4, IN5:=IN5);
  Ready := CollectInput.Finished;
  FeedNext := 1;
  IF Ready THEN
    Out := ((((((FALSE AND ((((Data[32] OR Data[11]) OR (Data[6] OR Data[33])) OR (Data[37] OR (NOT Data[33]))) OR (((Data[45] OR Data[22]) OR (NOT Data[44])) OR (NOT Data[47])))) OR (NOT (NOT Data[28]))) AND ((Data[24] XOR (((Data[3] AND ((((Data[19] AND Data[6]) AND ((Data[45] XOR Data[48]) XOR Data[8])) XOR (((NOT Data[33]) XOR (Data[26] AND Data[41])) XOR Data[48])) XOR ((((Data[48] XOR Data[4]) XOR Data[30]) XOR (Data[38] AND Data[7])) XOR (Data[2] AND Data[27])))) XOR ((((NOT Data[46]) AND (Data[25] AND Data[22])) OR Data[3]) AND Data[14])) XOR (((NOT ((Data[32] XOR Data[14]) XOR Data[46])) OR Data[41]) AND ((NOT (Data[32] OR Data[6])) AND (NOT (NOT Data[48])))))) XOR (NOT (((((Data[18] XOR Data[35]) XOR Data[47]) OR Data[25]) OR (((Data[1] OR Data[9]) XOR (Data[12] AND FALSE)) XOR TRUE)) AND (((Data[26] OR (Data[11] AND Data[20])) XOR Data[14]) XOR (NOT Data[41])))))) OR Data[15]) OR (NOT (NOT Data[18]))) OR Data[14]);
    OutReady := 1;
    CollectInput(RESET:=TRUE);
  END_IF;
END_PROGRAM

CONFIGURATION Config0
  RESOURCE Res0 ON PLC
    TASK task0(INTERVAL := T#20ms,PRIORITY := 0);
    PROGRAM instance0 WITH task0 : Boiler;
  END_RESOURCE
END_CONFIGURATION

(* ---- RND-EXPR_peens-since-gruel.st ---- *)
(*
This code implements a randomly grown symbolic expression:

xor(xor((!((((xor(xor(!(!(IN12 | IN12)), ((!(IN40)) | (IN7 & IN31)) | ((xor(xor(IN21, IN32), IN47)) & (IN27 | IN45))), !(!(!(IN26))))) | (xor(xor(IN6, ((IN4 & IN11) & (!(IN29))) | (!(!(IN9)))), (xor(xor(!(IN21), xor(xor(IN43, IN19), IN28)), IN32)) | true))) | (IN48 & ((((xor(xor(IN43, IN49), IN37)) | (xor(xor(IN48, IN12), IN29))) & (xor(xor(IN30, IN33 & IN29), IN3 & IN38))) & (IN36 & ((IN7 | IN5) & (!(IN22))))))) & IN15)) | IN23, IN44 | (!((IN10 & (xor(xor((!(!(IN9 & IN23))) & ((xor(xor(IN38 & IN15, xor(xor(IN1, IN44), IN41)), IN34)) | IN3), ((xor(xor(IN3 | IN10, xor(xor(IN26, IN48), IN11)), IN31 | IN9)) | (!(xor(xor(IN26, IN44), IN22)))) | IN7), (xor(xor(IN12, IN34), IN9 | IN19)) | IN37))) | (IN3 | IN16)))), xor(xor(true, IN41), xor(xor(xor(xor(IN27, ((xor(xor(!(IN6), xor(xor((xor(xor(IN12, IN43), IN35)) | (!(IN36)), xor(xor(IN34 | IN25, IN43 & IN12), !(IN16))), !(!(IN18)))), ((IN13 & IN1) | (IN4 | IN50)) & (!(xor(xor(IN12, IN13), IN23))))) & IN41) & (xor(xor((!((false | IN10) & (IN48 & IN31))) | (xor(xor(IN17, xor(xor(xor(xor(IN18, IN49), IN19), IN9), IN31)), (xor(xor(IN49, IN1), IN9)) & (xor(xor(IN9, IN31), IN42)))), ((IN4 | IN47) | IN2) | IN34), xor(xor(xor(xor((IN42 | IN4) | (IN12 | IN20), (!(IN8)) & (IN46 | IN24)), (IN8 | IN39) & true), (!(xor(xor(IN8, IN8), IN3))) & ((!(IN26)) & (IN31 | IN41))), !(IN32))))), !(((xor(xor((IN26 & IN24) | (IN3 | IN6), true & (true | IN44)), (xor(xor(IN36, IN8), IN39)) & (IN11 | IN3))) & ((!(IN10 | false)) & (xor(xor(IN22 & IN30, IN26), !(IN32))))) & IN8)), IN19), IN3 | ((((IN50 & (!(xor(xor(IN20, IN50), IN50)))) | ((xor(xor(IN41 | IN41, IN29 & IN48), IN9 & IN21)) | (xor(xor(xor(xor(IN11, IN46), IN46), IN5), !(IN50))))) | (!(xor(xor((IN11 & IN23) | (IN34 & IN20), (!(IN8)) & (xor(xor(IN37, true), IN12))), !(IN50 & IN14))))) | IN34))))

*)

FUNCTION_BLOCK F_CollectInput
  VAR_IN_OUT
      Data : ARRAY[1..50] OF BOOL;
  END_VAR
  VAR_INPUT
      TICK  : BOOL := 0;
      IN1   : BOOL := 0;
      IN2   : BOOL := 0;
      IN3   : BOOL := 0;
      IN4   : BOOL := 0;
      IN5   : BOOL := 0;
      RESET : BOOL := FALSE;
  END_VAR
  VAR_OUTPUT
      Finished : BOOL;
  END_VAR
  VAR
      j    : USINT := 1;
      tock : BOOL  := 0;
  END_VAR
  IF NOT RESET AND tock = NOT TICK THEN
      Data[j]   := IN1;
      Data[j+1] := IN2;
      Data[j+2] := IN3;
      Data[j+3] := IN4;
      Data[j+4] := IN5;
      j := j + 5;
      tock := TICK;
  ELSE
      j := 1;
      tock := 0;
  END_IF;
  Finished := (j > 50);
END_FUNCTION_BLOCK

PROGRAM Boiler
  VAR
    Data  : ARRAY[1..50] OF BOOL;
    Ready : BOOL;
    CollectInput : F_CollectInput;
  END_VAR
  VAR
    TICK     AT %IX1.0 : BOOL;
    IN1      AT %IX0.3 : BOOL;
    IN2      AT %IX0.4 : BOOL;
    IN3      AT %IX0.5 : BOOL;
    IN4      AT %IX0.6 : BOOL;
    IN5      AT %IX0.7 : BOOL;
    OutReady AT %QX0.0 : BOOL := FALSE;
    FeedNext AT %QX0.1 : BOOL := FALSE;
    Out      AT %QX0.2 : BOOL;
  END_VAR
  CollectInput(TICK:=TICK, IN1:=IN1, IN2:=IN2, IN3:=IN3, IN4:=IN4, IN5:=IN5);
  Ready := CollectInput.Finished;
  FeedNext := 1;
  IF Ready THEN
    Out := ((((NOT ((((((NOT (NOT (Data[12] OR Data[12]))) XOR (((NOT Data[40]) OR (Data[7] AND Data[31])) OR (((Data[21] XOR Data[32]) XOR Data[47]) AND (Data[27] OR Data[45])))) XOR (NOT (NOT (NOT Data[26])))) OR ((Data[6] XOR (((Data[4] AND Data[11]) AND (NOT Data[29])) OR (NOT (NOT Data[9])))) XOR ((((NOT Data[21]) XOR ((Data[43] XOR Data[19]) XOR Data[28])) XOR Data[32]) OR TRUE))) OR (Data[48] AND (((((Data[43] XOR Data[49]) XOR Data[37]) OR ((Data[48] XOR Data[12]) XOR Data[29])) AND ((Data[30] XOR (Data[33] AND Data[29])) XOR (Data[3] AND Data[38]))) AND (Data[36] AND ((Data[7] OR Data[5]) AND (NOT Data[22])))))) AND Data[15])) OR Data[23]) XOR (Data[44] OR (NOT ((Data[10] AND ((((NOT (NOT (Data[9] AND Data[23]))) AND ((((Data[38] AND Data[15]) XOR ((Data[1] XOR Data[44]) XOR Data[41])) XOR Data[34]) OR Data[3])) XOR (((((Data[3] OR Data[10]) XOR ((Data[26] XOR Data[48]) XOR Data[11])) XOR (Data[31] OR Data[9])) OR (NOT ((Data[26] XOR Data[44]) XOR Data[22]))) OR Data[7])) XOR (((Data[12] XOR Data[34]) XOR (Data[9] OR Data[19])) OR Data[37]))) OR (Data[3] OR Data[16]))))) XOR ((TRUE XOR Data[41]) XOR ((((Data[27] XOR (((((NOT Data[6]) XOR (((((Data[12] XOR Data[43]) XOR Data[35]) OR (NOT Data[36])) XOR (((Data[34] OR Data[25]) XOR (Data[43] AND Data[12])) XOR (NOT Data[16]))) XOR (NOT (NOT Data[18])))) XOR (((Data[13] AND Data[1]) OR (Data[4] OR Data[50])) AND (NOT ((Data[12] XOR Data[13]) XOR Data[23])))) AND Data[41]) AND ((((NOT ((FALSE OR Data[10]) AND (Data[48] AND Data[31]))) OR ((Data[17] XOR ((((Data[18] XOR Data[49]) XOR Data[19]) XOR Data[9]) XOR Data[31])) XOR (((Data[49] XOR Data[1]) XOR Data[9]) AND ((Data[9] XOR Data[31]) XOR Data[42])))) XOR (((Data[4] OR Data[47]) OR Data[2]) OR Data[34])) XOR ((((((Data[42] OR Data[4]) OR (Data[12] OR Data[20])) XOR ((NOT Data[8]) AND (Data[46] OR Data[24]))) XOR ((Data[8] OR Data[39]) AND TRUE)) XOR ((NOT ((Data[8] XOR Data[8]) XOR Data[3])) AND ((NOT Data[26]) AND (Data[31] OR Data[41])))) XOR (NOT Data[32]))))) XOR (NOT ((((((Data[26] AND Data[24]) OR (Data[3] OR Data[6])) XOR (TRUE AND (TRUE OR Data[44]))) XOR (((Data[36] XOR Data[8]) XOR Data[39]) AND (Data[11] OR Data[3]))) AND ((NOT (Data[10] OR FALSE)) AND (((Data[22] AND Data[30]) XOR Data[26]) XOR (NOT Data[32])))) AND Data[8]))) XOR Data[19]) XOR (Data[3] OR ((((Data[50] AND (NOT ((Data[20] XOR Data[50]) XOR Data[50]))) OR ((((Data[41] OR Data[41]) XOR (Data[29] AND Data[48])) XOR (Data[9] AND Data[21])) OR ((((Data[11] XOR Data[46]) XOR Data[46]) XOR Data[5]) XOR (NOT Data[50])))) OR (NOT ((((Data[11] AND Data[23]) OR (Data[34] AND Data[20])) XOR ((NOT Data[8]) AND ((Data[37] XOR TRUE) XOR Data[12]))) XOR (NOT (Data[50] AND Data[14]))))) OR Data[34])))));
    OutReady := 1;
    CollectInput(RESET:=TRUE);
  END_IF;
END_PROGRAM

CONFIGURATION Config0
  RESOURCE Res0 ON PLC
    TASK task0(INTERVAL := T#20ms,PRIORITY := 0);
    PROGRAM instance0 WITH task0 : Boiler;
  END_RESOURCE
END_CONFIGURATION

(* ---- RND-EXPR_pikes-stops-chill.st ---- *)
(*
This code implements a randomly grown symbolic expression:

!((IN16 & IN32) & ((xor(xor(xor(xor(IN24 | IN48, (((xor(xor(xor(xor(IN40, true), IN7), xor(xor(IN27, IN44), IN7)), IN6 | IN4)) & ((IN19 | IN14) & (IN40 & IN35))) & ((xor(xor(xor(xor(IN39, IN34), IN48), IN14), IN40)) | ((xor(xor(IN13, IN28), IN42)) & IN45))) & (!(((IN21 | IN2) & (xor(xor(IN10, IN37), IN37))) & (!(IN11))))), xor(xor(xor(xor(xor(xor(IN7, IN46), !(!(IN6))), !(!(IN40 & IN29))), ((IN46 | IN37) & IN8) & ((IN22 | IN10) & (!(IN45)))), IN18 & (((IN3 & IN7) | IN33) | (xor(xor(!(IN41), IN45), IN34 | IN4)))), (xor(xor(xor(xor(!(IN48), true), IN37), IN21), xor(xor(xor(xor(IN22, IN49), IN18), IN23 & IN36), xor(xor(IN50, IN46), IN46)))) & (!((IN47 & IN2) | (IN33 | IN12))))), !(IN49 | ((((!(IN38)) | (IN39 | IN16)) & ((IN6 | IN42) | IN24)) & (!((!(IN17)) & (true | IN18)))))), IN1)) & ((xor(xor(IN37, xor(xor(!(((IN10 | IN47) & (xor(xor(IN39, IN25), IN32))) & (xor(xor(!(IN11), IN27 | IN31), xor(xor(IN28, IN4), IN40)))), (xor(xor(!(IN50 & IN31), IN44), !(IN17 & IN29))) & ((!(IN47)) | ((!(IN16)) & (!(IN24))))), xor(xor(((!(IN19)) & (xor(xor(IN38, IN13), false))) & (xor(xor(IN15, IN34 | IN14), !(IN33))), xor(xor((xor(xor(IN39, IN24), IN44)) & IN42, (!(IN24)) & (xor(xor(IN23, IN12), IN20))), (xor(xor(false, IN3), IN48)) | (xor(xor(IN8, IN18), IN19)))), !((!(IN28)) | IN33)))), xor(xor(!(!(!(IN26 & false))), IN33), IN30 | ((IN48 | IN35) & (xor(xor(IN11 & IN12, IN29 | IN41), !(IN30))))))) & (xor(xor((IN8 & (!((IN8 | IN46) & IN22))) & (((!(IN29 & IN32)) | ((IN9 | IN45) & (!(IN24)))) | (((!(IN41)) | (xor(xor(IN1, IN37), IN29))) & ((IN13 | IN50) | (IN37 | IN11)))), !((xor(xor((IN17 | IN14) | (xor(xor(IN15, true), IN25)), !(xor(xor(IN2, IN26), IN23))), (IN37 | IN15) | (IN44 | IN22))) | ((xor(xor(xor(xor(IN23, IN31), IN33), IN39 | IN21), IN21)) | (!(!(IN19)))))), (!(((IN24 | false) | (xor(xor(IN17, IN50), IN9))) | (xor(xor(IN39 & IN35, IN19 & IN48), IN37 & IN25)))) | IN46)))))

*)

FUNCTION_BLOCK F_CollectInput
  VAR_IN_OUT
      Data : ARRAY[1..50] OF BOOL;
  END_VAR
  VAR_INPUT
      TICK  : BOOL := 0;
      IN1   : BOOL := 0;
      IN2   : BOOL := 0;
      IN3   : BOOL := 0;
      IN4   : BOOL := 0;
      IN5   : BOOL := 0;
      RESET : BOOL := FALSE;
  END_VAR
  VAR_OUTPUT
      Finished : BOOL;
  END_VAR
  VAR
      j    : USINT := 1;
      tock : BOOL  := 0;
  END_VAR
  IF NOT RESET AND tock = NOT TICK THEN
      Data[j]   := IN1;
      Data[j+1] := IN2;
      Data[j+2] := IN3;
      Data[j+3] := IN4;
      Data[j+4] := IN5;
      j := j + 5;
      tock := TICK;
  ELSE
      j := 1;
      tock := 0;
  END_IF;
  Finished := (j > 50);
END_FUNCTION_BLOCK

PROGRAM Boiler
  VAR
    Data  : ARRAY[1..50] OF BOOL;
    Ready : BOOL;
    CollectInput : F_CollectInput;
  END_VAR
  VAR
    TICK     AT %IX1.0 : BOOL;
    IN1      AT %IX0.3 : BOOL;
    IN2      AT %IX0.4 : BOOL;
    IN3      AT %IX0.5 : BOOL;
    IN4      AT %IX0.6 : BOOL;
    IN5      AT %IX0.7 : BOOL;
    OutReady AT %QX0.0 : BOOL := FALSE;
    FeedNext AT %QX0.1 : BOOL := FALSE;
    Out      AT %QX0.2 : BOOL;
  END_VAR
  CollectInput(TICK:=TICK, IN1:=IN1, IN2:=IN2, IN3:=IN3, IN4:=IN4, IN5:=IN5);
  Ready := CollectInput.Finished;
  FeedNext := 1;
  IF Ready THEN
    Out := (NOT ((Data[16] AND Data[32]) AND ((((((Data[24] OR Data[48]) XOR (((((((Data[40] XOR TRUE) XOR Data[7]) XOR ((Data[27] XOR Data[44]) XOR Data[7])) XOR (Data[6] OR Data[4])) AND ((Data[19] OR Data[14]) AND (Data[40] AND Data[35]))) AND (((((Data[39] XOR Data[34]) XOR Data[48]) XOR Data[14]) XOR Data[40]) OR (((Data[13] XOR Data[28]) XOR Data[42]) AND Data[45]))) AND (NOT (((Data[21] OR Data[2]) AND ((Data[10] XOR Data[37]) XOR Data[37])) AND (NOT Data[11]))))) XOR ((((((Data[7] XOR Data[46]) XOR (NOT (NOT Data[6]))) XOR (NOT (NOT (Data[40] AND Data[29])))) XOR (((Data[46] OR Data[37]) AND Data[8]) AND ((Data[22] OR Data[10]) AND (NOT Data[45])))) XOR (Data[18] AND (((Data[3] AND Data[7]) OR Data[33]) OR (((NOT Data[41]) XOR Data[45]) XOR (Data[34] OR Data[4]))))) XOR ((((((NOT Data[48]) XOR TRUE) XOR Data[37]) XOR Data[21]) XOR ((((Data[22] XOR Data[49]) XOR Data[18]) XOR (Data[23] AND Data[36])) XOR ((Data[50] XOR Data[46]) XOR Data[46]))) AND (NOT ((Data[47] AND Data[2]) OR (Data[33] OR Data[12])))))) XOR (NOT (Data[49] OR ((((NOT Data[38]) OR (Data[39] OR Data[16])) AND ((Data[6] OR Data[42]) OR Data[24])) AND (NOT ((NOT Data[17]) AND (TRUE OR Data[18]))))))) XOR Data[1]) AND (((Data[37] XOR (((NOT (((Data[10] OR Data[47]) AND ((Data[39] XOR Data[25]) XOR Data[32])) AND (((NOT Data[11]) XOR (Data[27] OR Data[31])) XOR ((Data[28] XOR Data[4]) XOR Data[40])))) XOR ((((NOT (Data[50] AND Data[31])) XOR Data[44]) XOR (NOT (Data[17] AND Data[29]))) AND ((NOT Data[47]) OR ((NOT Data[16]) AND (NOT Data[24]))))) XOR (((((NOT Data[19]) AND ((Data[38] XOR Data[13]) XOR FALSE)) AND ((Data[15] XOR (Data[34] OR Data[14])) XOR (NOT Data[33]))) XOR (((((Data[39] XOR Data[24]) XOR Data[44]) AND Data[42]) XOR ((NOT Data[24]) AND ((Data[23] XOR Data[12]) XOR Data[20]))) XOR (((FALSE XOR Data[3]) XOR Data[48]) OR ((Data[8] XOR Data[18]) XOR Data[19])))) XOR (NOT ((NOT Data[28]) OR Data[33]))))) XOR (((NOT (NOT (NOT (Data[26] AND FALSE)))) XOR Data[33]) XOR (Data[30] OR ((Data[48] OR Data[35]) AND (((Data[11] AND Data[12]) XOR (Data[29] OR Data[41])) XOR (NOT Data[30])))))) AND ((((Data[8] AND (NOT ((Data[8] OR Data[46]) AND Data[22]))) AND (((NOT (Data[29] AND Data[32])) OR ((Data[9] OR Data[45]) AND (NOT Data[24]))) OR (((NOT Data[41]) OR ((Data[1] XOR Data[37]) XOR Data[29])) AND ((Data[13] OR Data[50]) OR (Data[37] OR Data[11]))))) XOR (NOT (((((Data[17] OR Data[14]) OR ((Data[15] XOR TRUE) XOR Data[25])) XOR (NOT ((Data[2] XOR Data[26]) XOR Data[23]))) XOR ((Data[37] OR Data[15]) OR (Data[44] OR Data[22]))) OR (((((Data[23] XOR Data[31]) XOR Data[33]) XOR (Data[39] OR Data[21])) XOR Data[21]) OR (NOT (NOT Data[19])))))) XOR ((NOT (((Data[24] OR FALSE) OR ((Data[17] XOR Data[50]) XOR Data[9])) OR (((Data[39] AND Data[35]) XOR (Data[19] AND Data[48])) XOR (Data[37] AND Data[25])))) OR Data[46]))))));
    OutReady := 1;
    CollectInput(RESET:=TRUE);
  END_IF;
END_PROGRAM

CONFIGURATION Config0
  RESOURCE Res0 ON PLC
    TASK task0(INTERVAL := T#20ms,PRIORITY := 0);
    PROGRAM instance0 WITH task0 : Boiler;
  END_RESOURCE
END_CONFIGURATION

(* ---- RND-EXPR_prods-erase-cores.st ---- *)
(*
This code implements a randomly grown symbolic expression:

xor(xor(true, xor(xor(IN39, (IN10 | (((xor(xor((!(IN45 | IN10)) | (xor(xor(IN33, IN25), xor(xor(IN10, IN32), IN30))), true & IN23), ((IN2 | IN2) & (xor(xor(IN34, IN12), IN29))) | ((IN49 | IN18) & (!(IN31))))) & ((((IN11 | IN46) & (IN6 & IN34)) | (!(IN49 | IN9))) | IN24)) | IN19)) | (xor(xor((xor(xor(!(!(!(!(IN24)))), IN24), (IN47 | (!(IN23))) | ((xor(xor(IN22, IN43 & IN35), !(IN43))) & IN24))) | ((xor(xor(IN7 | (!(IN47 & IN26)), !(!(IN40))), !((xor(xor(IN29, IN40), IN14)) & (xor(xor(IN41, IN9), IN5))))) | ((xor(xor(xor(xor(IN29 | IN41, IN41 | IN39), xor(xor(IN34, IN15), IN12)), xor(xor(xor(xor(IN14, IN40), IN45), !(IN43)), IN47 | IN20)), (xor(xor(IN32, IN12), IN48)) | (xor(xor(IN7, IN6), IN12)))) | ((xor(xor(false | IN50, IN3 | IN49), xor(xor(IN48, IN10), IN47))) | ((xor(xor(IN1, IN39), IN16)) | (!(IN23)))))), xor(xor(!((((xor(xor(IN1, IN3), IN11)) | (IN48 & IN36)) | ((IN44 | IN11) & (IN23 & IN15))) | ((!(IN6 & false)) | (!(IN22 & IN2)))), IN8), ((((!(IN41)) & (IN48 & IN48)) | (xor(xor(xor(xor(IN10, IN25), IN34), xor(xor(IN36, true), IN11)), IN40 & IN26))) & (!(IN46))) | (xor(xor(!(!(IN5)), IN2), xor(xor(xor(xor(xor(xor(IN7, IN26), IN48), IN40), IN50), IN7), (IN14 | IN3) & (!(IN25))))))), IN6))), IN17)), (!(IN46 | IN27)) | ((xor(xor(xor(xor((xor(xor(!((IN17 & IN1) & (IN39 | IN43)), IN36), IN6)) & (!(IN10 | (IN12 | (xor(xor(IN14, IN1), IN33))))), xor(xor(xor(xor(!((IN45 & IN11) & IN26), IN46), xor(xor(IN4 & (IN25 & IN13), (!(IN13)) & (xor(xor(IN3, IN35), IN38))), xor(xor(IN8, xor(xor(IN28, IN15), IN7)), !(IN39)))), xor(xor(IN29 & ((!(IN29)) | (IN42 | IN32)), !(IN36)), (IN43 | (IN27 | IN37)) | ((IN4 | IN3) & (xor(xor(IN30, IN14), IN13))))), xor(xor(xor(xor(IN17, IN48), IN45), IN2), ((IN23 & IN16) & false) | (xor(xor(IN14, IN25 | IN47), xor(xor(IN50, IN26), IN42)))))), !(!(xor(xor((IN16 & false) | (IN22 & IN30), (IN12 & true) & (!(IN32))), (IN5 | IN37) | IN45)))), xor(xor(IN36, (xor(xor(!(!(!(IN7))), !(IN33)), !(xor(xor(IN24 & IN22, IN27 | IN13), true & IN24)))) | ((((!(IN50)) & IN15) & (xor(xor(xor(xor(IN37, IN21), IN23), !(IN49)), !(IN31)))) | (xor(xor(IN7 & (!(IN31)), IN28), (IN47 | IN33) & IN3)))), ((!(xor(xor(xor(xor(IN23, IN29), IN9), !(IN29)), IN44))) | (((!(IN8)) | IN50) & ((IN7 | IN10) | (IN30 & IN33)))) | (xor(xor(((IN44 | IN39) | (IN50 & IN42)) & (xor(xor(IN10 & IN47, IN19), IN34 | IN26)), xor(xor(IN19, !(IN15 & IN12)), !(!(IN7)))), !((xor(xor(IN41, IN13), IN29)) & IN2))))), IN44)) | (xor(xor(IN20 & (IN42 | ((!((IN24 | IN45) | (IN37 | IN7))) & ((xor(xor(IN2 | false, xor(xor(IN49, IN27), IN44)), IN31)) | IN16))), IN39 | (!(xor(xor(IN10, ((IN50 | IN21) | (IN23 | IN29)) & ((IN32 & IN12) & (IN43 & IN21))), xor(xor(xor(xor(IN50 | false, xor(xor(IN45, IN30), IN29)), IN27 & IN7), !(IN42 | IN35)), (IN18 & IN8) | (IN11 | IN5)))))), xor(xor(((!(!(!(IN24)))) | IN42) | IN35, xor(xor((!((xor(xor(IN11, IN48), true)) | (IN3 | IN48))) & ((IN19 & (IN49 | IN38)) | (xor(xor(!(IN35), !(IN20)), IN2 | IN33))), IN14), ((!(!(IN36))) | (true & (xor(xor(IN36, IN34), IN35)))) & (((IN28 & IN27) & (IN6 & IN47)) | (IN30 | (IN43 & IN16))))), xor(xor((IN20 & ((IN10 | IN10) & IN47)) | IN16, ((xor(xor(IN8 | IN1, IN43), !(IN7))) & ((xor(xor(IN8, IN28), IN43)) | IN9)) & IN14), ((!(!(IN47))) | ((!(IN50)) & (IN27 & IN46))) & (xor(xor((IN14 & IN40) | (IN17 | IN2), xor(xor(IN20 | IN31, IN28 & IN19), IN50 & IN40)), (IN4 | IN35) & (xor(xor(IN40, IN16), IN32))))))))))

*)

FUNCTION_BLOCK F_CollectInput
  VAR_IN_OUT
      Data : ARRAY[1..50] OF BOOL;
  END_VAR
  VAR_INPUT
      TICK  : BOOL := 0;
      IN1   : BOOL := 0;
      IN2   : BOOL := 0;
      IN3   : BOOL := 0;
      IN4   : BOOL := 0;
      IN5   : BOOL := 0;
      RESET : BOOL := FALSE;
  END_VAR
  VAR_OUTPUT
      Finished : BOOL;
  END_VAR
  VAR
      j    : USINT := 1;
      tock : BOOL  := 0;
  END_VAR
  IF NOT RESET AND tock = NOT TICK THEN
      Data[j]   := IN1;
      Data[j+1] := IN2;
      Data[j+2] := IN3;
      Data[j+3] := IN4;
      Data[j+4] := IN5;
      j := j + 5;
      tock := TICK;
  ELSE
      j := 1;
      tock := 0;
  END_IF;
  Finished := (j > 50);
END_FUNCTION_BLOCK

PROGRAM Boiler
  VAR
    Data  : ARRAY[1..50] OF BOOL;
    Ready : BOOL;
    CollectInput : F_CollectInput;
  END_VAR
  VAR
    TICK     AT %IX1.0 : BOOL;
    IN1      AT %IX0.3 : BOOL;
    IN2      AT %IX0.4 : BOOL;
    IN3      AT %IX0.5 : BOOL;
    IN4      AT %IX0.6 : BOOL;
    IN5      AT %IX0.7 : BOOL;
    OutReady AT %QX0.0 : BOOL := FALSE;
    FeedNext AT %QX0.1 : BOOL := FALSE;
    Out      AT %QX0.2 : BOOL;
  END_VAR
  CollectInput(TICK:=TICK, IN1:=IN1, IN2:=IN2, IN3:=IN3, IN4:=IN4, IN5:=IN5);
  Ready := CollectInput.Finished;
  FeedNext := 1;
  IF Ready THEN
    Out := ((TRUE XOR ((Data[39] XOR ((Data[10] OR ((((((NOT (Data[45] OR Data[10])) OR ((Data[33] XOR Data[25]) XOR ((Data[10] XOR Data[32]) XOR Data[30]))) XOR (TRUE AND Data[23])) XOR (((Data[2] OR Data[2]) AND ((Data[34] XOR Data[12]) XOR Data[29])) OR ((Data[49] OR Data[18]) AND (NOT Data[31])))) AND ((((Data[11] OR Data[46]) AND (Data[6] AND Data[34])) OR (NOT (Data[49] OR Data[9]))) OR Data[24])) OR Data[19])) OR ((((((NOT (NOT (NOT (NOT Data[24])))) XOR Data[24]) XOR ((Data[47] OR (NOT Data[23])) OR (((Data[22] XOR (Data[43] AND Data[35])) XOR (NOT Data[43])) AND Data[24]))) OR ((((Data[7] OR (NOT (Data[47] AND Data[26]))) XOR (NOT (NOT Data[40]))) XOR (NOT (((Data[29] XOR Data[40]) XOR Data[14]) AND ((Data[41] XOR Data[9]) XOR Data[5])))) OR ((((((Data[29] OR Data[41]) XOR (Data[41] OR Data[39])) XOR ((Data[34] XOR Data[15]) XOR Data[12])) XOR ((((Data[14] XOR Data[40]) XOR Data[45]) XOR (NOT Data[43])) XOR (Data[47] OR Data[20]))) XOR (((Data[32] XOR Data[12]) XOR Data[48]) OR ((Data[7] XOR Data[6]) XOR Data[12]))) OR ((((FALSE OR Data[50]) XOR (Data[3] OR Data[49])) XOR ((Data[48] XOR Data[10]) XOR Data[47])) OR (((Data[1] XOR Data[39]) XOR Data[16]) OR (NOT Data[23])))))) XOR (((NOT (((((Data[1] XOR Data[3]) XOR Data[11]) OR (Data[48] AND Data[36])) OR ((Data[44] OR Data[11]) AND (Data[23] AND Data[15]))) OR ((NOT (Data[6] AND FALSE)) OR (NOT (Data[22] AND Data[2]))))) XOR Data[8]) XOR (((((NOT Data[41]) AND (Data[48] AND Data[48])) OR ((((Data[10] XOR Data[25]) XOR Data[34]) XOR ((Data[36] XOR TRUE) XOR Data[11])) XOR (Data[40] AND Data[26]))) AND (NOT Data[46])) OR (((NOT (NOT Data[5])) XOR Data[2]) XOR ((((((Data[7] XOR Data[26]) XOR Data[48]) XOR Data[40]) XOR Data[50]) XOR Data[7]) XOR ((Data[14] OR Data[3]) AND (NOT Data[25]))))))) XOR Data[6]))) XOR Data[17])) XOR ((NOT (Data[46] OR Data[27])) OR (((((((((NOT ((Data[17] AND Data[1]) AND (Data[39] OR Data[43]))) XOR Data[36]) XOR Data[6]) AND (NOT (Data[10] OR (Data[12] OR ((Data[14] XOR Data[1]) XOR Data[33]))))) XOR (((((NOT ((Data[45] AND Data[11]) AND Data[26])) XOR Data[46]) XOR (((Data[4] AND (Data[25] AND Data[13])) XOR ((NOT Data[13]) AND ((Data[3] XOR Data[35]) XOR Data[38]))) XOR ((Data[8] XOR ((Data[28] XOR Data[15]) XOR Data[7])) XOR (NOT Data[39])))) XOR (((Data[29] AND ((NOT Data[29]) OR (Data[42] OR Data[32]))) XOR (NOT Data[36])) XOR ((Data[43] OR (Data[27] OR Data[37])) OR ((Data[4] OR Data[3]) AND ((Data[30] XOR Data[14]) XOR Data[13]))))) XOR ((((Data[17] XOR Data[48]) XOR Data[45]) XOR Data[2]) XOR (((Data[23] AND Data[16]) AND FALSE) OR ((Data[14] XOR (Data[25] OR Data[47])) XOR ((Data[50] XOR Data[26]) XOR Data[42])))))) XOR (NOT (NOT ((((Data[16] AND FALSE) OR (Data[22] AND Data[30])) XOR ((Data[12] AND TRUE) AND (NOT Data[32]))) XOR ((Data[5] OR Data[37]) OR Data[45]))))) XOR ((Data[36] XOR ((((NOT (NOT (NOT Data[7]))) XOR (NOT Data[33])) XOR (NOT (((Data[24] AND Data[22]) XOR (Data[27] OR Data[13])) XOR (TRUE AND Data[24])))) OR ((((NOT Data[50]) AND Data[15]) AND ((((Data[37] XOR Data[21]) XOR Data[23]) XOR (NOT Data[49])) XOR (NOT Data[31]))) OR (((Data[7] AND (NOT Data[31])) XOR Data[28]) XOR ((Data[47] OR Data[33]) AND Data[3]))))) XOR (((NOT ((((Data[23] XOR Data[29]) XOR Data[9]) XOR (NOT Data[29])) XOR Data[44])) OR (((NOT Data[8]) OR Data[50]) AND ((Data[7] OR Data[10]) OR (Data[30] AND Data[33])))) OR (((((Data[44] OR Data[39]) OR (Data[50] AND Data[42])) AND (((Data[10] AND Data[47]) XOR Data[19]) XOR (Data[34] OR Data[26]))) XOR ((Data[19] XOR (NOT (Data[15] AND Data[12]))) XOR (NOT (NOT Data[7])))) XOR (NOT (((Data[41] XOR Data[13]) XOR Data[29]) AND Data[2])))))) XOR Data[44]) OR (((Data[20] AND (Data[42] OR ((NOT ((Data[24] OR Data[45]) OR (Data[37] OR Data[7]))) AND ((((Data[2] OR FALSE) XOR ((Data[49] XOR Data[27]) XOR Data[44])) XOR Data[31]) OR Data[16])))) XOR (Data[39] OR (NOT ((Data[10] XOR (((Data[50] OR Data[21]) OR (Data[23] OR Data[29])) AND ((Data[32] AND Data[12]) AND (Data[43] AND Data[21])))) XOR (((((Data[50] OR FALSE) XOR ((Data[45] XOR Data[30]) XOR Data[29])) XOR (Data[27] AND Data[7])) XOR (NOT (Data[42] OR Data[35]))) XOR ((Data[18] AND Data[8]) OR (Data[11] OR Data[5]))))))) XOR (((((NOT (NOT (NOT Data[24]))) OR Data[42]) OR Data[35]) XOR ((((NOT (((Data[11] XOR Data[48]) XOR TRUE) OR (Data[3] OR Data[48]))) AND ((Data[19] AND (Data[49] OR Data[38])) OR (((NOT Data[35]) XOR (NOT Data[20])) XOR (Data[2] OR Data[33])))) XOR Data[14]) XOR (((NOT (NOT Data[36])) OR (TRUE AND ((Data[36] XOR Data[34]) XOR Data[35]))) AND (((Data[28] AND Data[27]) AND (Data[6] AND Data[47])) OR (Data[30] OR (Data[43] AND Data[16])))))) XOR ((((Data[20] AND ((Data[10] OR Data[10]) AND Data[47])) OR Data[16]) XOR (((((Data[8] OR Data[1]) XOR Data[43]) XOR (NOT Data[7])) AND (((Data[8] XOR Data[28]) XOR Data[43]) OR Data[9])) AND Data[14])) XOR (((NOT (NOT Data[47])) OR ((NOT Data[50]) AND (Data[27] AND Data[46]))) AND ((((Data[14] AND Data[40]) OR (Data[17] OR Data[2])) XOR (((Data[20] OR Data[31]) XOR (Data[28] AND Data[19])) XOR (Data[50] AND Data[40]))) XOR ((Data[4] OR Data[35]) AND ((Data[40] XOR Data[16]) XOR Data[32]))))))))));
    OutReady := 1;
    CollectInput(RESET:=TRUE);
  END_IF;
END_PROGRAM

CONFIGURATION Config0
  RESOURCE Res0 ON PLC
    TASK task0(INTERVAL := T#20ms,PRIORITY := 0);
    PROGRAM instance0 WITH task0 : Boiler;
  END_RESOURCE
END_CONFIGURATION

(* ---- RND-EXPR_purrs-djinn-ritzy.st ---- *)
(*
This code implements a randomly grown symbolic expression:

((!((IN27 & (!(((IN20 & (xor(xor(IN19, IN43), IN36))) | (!(xor(xor(IN23, IN22), IN14)))) & (!(IN16))))) | (((!(xor(xor(!(IN30 | IN14), !(IN23 | IN26)), !(xor(xor(IN44, IN12), IN19))))) & (!(IN5))) & IN9))) | ((IN46 & (!(!(IN11)))) & (xor(xor(IN5 & (xor(xor(!(!((IN38 | IN42) & (xor(xor(IN48, IN50), IN13)))), (xor(xor(IN49, IN50 | (!(IN24))), IN31)) | ((IN37 | (IN48 | IN34)) & ((IN35 | IN16) | (IN17 | IN43)))), IN13 | IN10)), (IN33 & ((!(IN17)) & (IN34 & IN48))) | IN32), IN5 & (IN20 | (xor(xor(IN25, IN24 | (IN15 & (!(IN8)))), IN27))))))) | ((!((xor(xor(!(IN27), IN41), xor(xor(xor(xor(IN26, (xor(xor(IN36 | IN34, xor(xor(IN21, IN29), IN42)), IN4)) | ((xor(xor(IN32, IN17), IN42)) & (IN8 & IN26))), (IN38 | (!(IN47))) & ((xor(xor(IN50, IN16), IN26)) & IN16)), (!((IN33 & IN46) | (IN1 | IN18))) & ((xor(xor(IN27 | IN36, IN18 & IN42), xor(xor(IN4, IN42), IN39))) & (IN45 & (xor(xor(IN42, IN15), IN42))))), !((!(xor(xor(IN47, IN15), IN19))) & IN30)))) & (!(xor(xor(IN2, (!(xor(xor(IN41, IN14 | IN24), xor(xor(IN45, IN37), IN19)))) & IN41), IN15 & (!((IN25 | true) & (IN41 | IN32)))))))) | (IN34 & (!((xor(xor(true, !(xor(xor(xor(xor(xor(xor(IN39, IN9), IN41), xor(xor(IN37, IN26), IN31)), xor(xor(IN21, IN3), IN24)), !(IN23 & IN19)), !(!(IN14))))), (((IN22 & false) | (!(IN12))) | (IN38 & (IN4 & IN30))) | ((xor(xor(!(IN27), IN31 & IN36), !(IN19))) & (!(!(IN1)))))) & (!(IN13))))))

*)

FUNCTION_BLOCK F_CollectInput
  VAR_IN_OUT
      Data : ARRAY[1..50] OF BOOL;
  END_VAR
  VAR_INPUT
      TICK  : BOOL := 0;
      IN1   : BOOL := 0;
      IN2   : BOOL := 0;
      IN3   : BOOL := 0;
      IN4   : BOOL := 0;
      IN5   : BOOL := 0;
      RESET : BOOL := FALSE;
  END_VAR
  VAR_OUTPUT
      Finished : BOOL;
  END_VAR
  VAR
      j    : USINT := 1;
      tock : BOOL  := 0;
  END_VAR
  IF NOT RESET AND tock = NOT TICK THEN
      Data[j]   := IN1;
      Data[j+1] := IN2;
      Data[j+2] := IN3;
      Data[j+3] := IN4;
      Data[j+4] := IN5;
      j := j + 5;
      tock := TICK;
  ELSE
      j := 1;
      tock := 0;
  END_IF;
  Finished := (j > 50);
END_FUNCTION_BLOCK

PROGRAM Boiler
  VAR
    Data  : ARRAY[1..50] OF BOOL;
    Ready : BOOL;
    CollectInput : F_CollectInput;
  END_VAR
  VAR
    TICK     AT %IX1.0 : BOOL;
    IN1      AT %IX0.3 : BOOL;
    IN2      AT %IX0.4 : BOOL;
    IN3      AT %IX0.5 : BOOL;
    IN4      AT %IX0.6 : BOOL;
    IN5      AT %IX0.7 : BOOL;
    OutReady AT %QX0.0 : BOOL := FALSE;
    FeedNext AT %QX0.1 : BOOL := FALSE;
    Out      AT %QX0.2 : BOOL;
  END_VAR
  CollectInput(TICK:=TICK, IN1:=IN1, IN2:=IN2, IN3:=IN3, IN4:=IN4, IN5:=IN5);
  Ready := CollectInput.Finished;
  FeedNext := 1;
  IF Ready THEN
    Out := (((NOT ((Data[27] AND (NOT (((Data[20] AND ((Data[19] XOR Data[43]) XOR Data[36])) OR (NOT ((Data[23] XOR Data[22]) XOR Data[14]))) AND (NOT Data[16])))) OR (((NOT (((NOT (Data[30] OR Data[14])) XOR (NOT (Data[23] OR Data[26]))) XOR (NOT ((Data[44] XOR Data[12]) XOR Data[19])))) AND (NOT Data[5])) AND Data[9]))) OR ((Data[46] AND (NOT (NOT Data[11]))) AND (((Data[5] AND (((NOT (NOT ((Data[38] OR Data[42]) AND ((Data[48] XOR Data[50]) XOR Data[13])))) XOR (((Data[49] XOR (Data[50] OR (NOT Data[24]))) XOR Data[31]) OR ((Data[37] OR (Data[48] OR Data[34])) AND ((Data[35] OR Data[16]) OR (Data[17] OR Data[43]))))) XOR (Data[13] OR Data[10]))) XOR ((Data[33] AND ((NOT Data[17]) AND (Data[34] AND Data[48]))) OR Data[32])) XOR (Data[5] AND (Data[20] OR ((Data[25] XOR (Data[24] OR (Data[15] AND (NOT Data[8])))) XOR Data[27])))))) OR ((NOT ((((NOT Data[27]) XOR Data[41]) XOR ((((Data[26] XOR ((((Data[36] OR Data[34]) XOR ((Data[21] XOR Data[29]) XOR Data[42])) XOR Data[4]) OR (((Data[32] XOR Data[17]) XOR Data[42]) AND (Data[8] AND Data[26])))) XOR ((Data[38] OR (NOT Data[47])) AND (((Data[50] XOR Data[16]) XOR Data[26]) AND Data[16]))) XOR ((NOT ((Data[33] AND Data[46]) OR (Data[1] OR Data[18]))) AND ((((Data[27] OR Data[36]) XOR (Data[18] AND Data[42])) XOR ((Data[4] XOR Data[42]) XOR Data[39])) AND (Data[45] AND ((Data[42] XOR Data[15]) XOR Data[42]))))) XOR (NOT ((NOT ((Data[47] XOR Data[15]) XOR Data[19])) AND Data[30])))) AND (NOT ((Data[2] XOR ((NOT ((Data[41] XOR (Data[14] OR Data[24])) XOR ((Data[45] XOR Data[37]) XOR Data[19]))) AND Data[41])) XOR (Data[15] AND (NOT ((Data[25] OR TRUE) AND (Data[41] OR Data[32])))))))) OR (Data[34] AND (NOT (((TRUE XOR (NOT ((((((Data[39] XOR Data[9]) XOR Data[41]) XOR ((Data[37] XOR Data[26]) XOR Data[31])) XOR ((Data[21] XOR Data[3]) XOR Data[24])) XOR (NOT (Data[23] AND Data[19]))) XOR (NOT (NOT Data[14]))))) XOR ((((Data[22] AND FALSE) OR (NOT Data[12])) OR (Data[38] AND (Data[4] AND Data[30]))) OR ((((NOT Data[27]) XOR (Data[31] AND Data[36])) XOR (NOT Data[19])) AND (NOT (NOT Data[1]))))) AND (NOT Data[13]))))));
    OutReady := 1;
    CollectInput(RESET:=TRUE);
  END_IF;
END_PROGRAM

CONFIGURATION Config0
  RESOURCE Res0 ON PLC
    TASK task0(INTERVAL := T#20ms,PRIORITY := 0);
    PROGRAM instance0 WITH task0 : Boiler;
  END_RESOURCE
END_CONFIGURATION

(* ---- RND-EXPR_races-touts-gaunt.st ---- *)
(*
This code implements a randomly grown symbolic expression:

(xor(xor((IN23 & IN50) | true, !(xor(xor(xor(xor(IN2 & ((xor(xor(IN36, IN7 | IN13), (!(IN18)) & (!(IN35)))) | (xor(xor((IN26 & IN39) & (xor(xor(IN30, IN3), IN8)), xor(xor(xor(xor(IN44, IN21), IN35), IN13 | IN29), xor(xor(IN6, IN46), IN32))), (!(IN27)) | (IN49 | IN27)))), !(IN28 | IN36)), IN31), (xor(xor(xor(xor(xor(xor(xor(xor(xor(xor(IN26, IN14), IN11), xor(xor(IN42, IN50), IN34)), IN29), !(IN42)), IN17), IN33), xor(xor(IN2 & (IN40 & IN9), IN26 & (IN23 | IN38)), IN10)), ((IN23 | (xor(xor(IN49, IN18), IN18))) | (xor(xor(xor(xor(IN10, IN38), IN17), IN31 & IN19), IN50 | IN39))) | (!(xor(xor(!(IN15), xor(xor(IN10, IN30), IN41)), IN17)))), IN41)) & (!(xor(xor(IN23, IN34 & (xor(xor(IN7 | IN19, IN31 & IN35), !(IN42)))), (!(IN36 & IN35)) & ((!(IN6)) & (IN9 | IN17)))))), IN6))), (!(((((!(IN6)) | ((IN19 & IN9) | (IN47 | IN24))) | (((!(IN43)) | (xor(xor(IN29, IN49), IN49))) | IN34)) | IN19) | (xor(xor(!(xor(xor(IN21, !(IN35)), !(!(IN7)))), IN31), (false & ((IN27 | IN44) | IN9)) | (((IN16 | IN28) | (IN33 | IN40)) | (!(IN34))))))) & ((!(IN38 | (IN30 | (xor(xor((xor(xor(IN31, IN2), IN4)) | (IN29 & IN7), !(xor(xor(IN7, false), IN43))), (xor(xor(IN23, IN28), IN27)) & IN20))))) | (((!((xor(xor(IN22, xor(xor(IN45, IN6), IN27)), IN21)) | (IN36 & (IN47 & IN2)))) & ((((IN12 | IN27) & (IN27 & IN26)) & (IN6 | (IN3 & IN10))) & (((IN44 | IN37) | (IN17 | IN19)) | (xor(xor(IN11 & IN29, IN2), !(IN40)))))) & (((((xor(xor(IN50, IN4), IN25)) | (!(IN12))) | (xor(xor(IN13 | IN7, IN10 & IN39), IN47))) | true) | (xor(xor(xor(xor(xor(xor(IN27 | IN11, IN42 & IN28), IN19 | IN24), false), (IN28 | IN32) | (!(IN49))), !(IN50)), (!(xor(xor(IN40, IN5), IN7))) & (!(IN40))))))))) & ((xor(xor(!((!(((!(xor(xor(IN34, IN33), IN17))) | ((IN20 & IN38) & (IN39 & IN6))) & (IN12 & (!(xor(xor(IN9, IN5), IN8)))))) & (xor(xor(xor(xor(IN11, !(xor(xor(IN50 | IN26, !(IN33)), IN14))), IN32), ((!(IN27 | IN20)) & (xor(xor(!(IN38), IN14 | IN18), IN30 & IN44))) & (!((IN45 & IN35) & (IN28 & IN49)))), xor(xor(IN8, (!(xor(xor(IN48, IN20), IN10))) | IN9), (!(!(IN28))) & (xor(xor(IN17 & IN28, !(IN35)), IN9 | IN18)))))), IN41 | (!(xor(xor((!((IN5 & IN1) | (xor(xor(IN50, IN32), IN38)))) & true, xor(xor(xor(xor(!(xor(xor(IN11, IN43), IN38)), xor(xor(xor(xor(IN49, IN30), IN35), IN34 & IN33), IN19 | IN27)), (IN9 & IN18) & (xor(xor(false, IN7), IN40))), (xor(xor(IN15 | IN48, IN45), !(IN47))) | ((!(IN44)) & (!(IN21)))), xor(xor((IN15 | IN44) & (!(IN2)), (IN10 | IN4) | (!(IN14))), false))), IN8)))), IN12)) & (xor(xor(xor(xor((xor(xor(IN28, !(xor(xor(IN36, IN8 & (IN6 | IN28)), xor(xor(xor(xor(IN44, IN8), IN44), IN16 | IN15), IN36 | IN22)))), IN40)) & (xor(xor(xor(xor(IN8, ((IN48 | IN38) | (xor(xor(IN40, IN46), IN32))) | ((xor(xor(IN15, IN16), IN46)) | IN25)), !(!(!(IN17)))), xor(xor(((IN1 | IN16) & (IN2 | IN15)) & (!(IN19)), ((IN42 | IN44) | IN35) & (!(IN48 | IN35))), IN3)), xor(xor(((IN9 & IN26) & (xor(xor(IN1, IN30), IN16))) & (IN9 | (xor(xor(IN4, IN44), IN15))), (!(xor(xor(IN47, IN5), IN41))) & (IN18 | (xor(xor(IN9, IN45), IN23)))), !(IN32)))), ((xor(xor(!(IN27), IN9), (xor(xor(IN16, IN41 | IN36), IN41)) | (xor(xor(IN48, IN22), IN25 & IN36)))) | (!(IN46 & ((xor(xor(IN16, IN48), IN39)) | (xor(xor(IN15, true), IN12)))))) | IN44), IN48 & ((!(!((IN27 & IN33) & (IN33 & IN39)))) | (IN19 & IN41))), !(IN40)), !((xor(xor(xor(xor(xor(xor(xor(xor(IN30 | IN38, xor(xor(IN39, IN19), IN33)), IN40 | IN13), IN44), (!(IN26)) & IN23), ((IN16 | IN48) & IN22) | (IN23 & (IN1 & IN3))), IN8), (!((IN43 & IN11) & IN33)) & IN16), (!((xor(xor(IN47, IN34), IN37)) | (!(IN19)))) | ((!(IN27)) & ((xor(xor(IN3, IN37), IN48)) | IN22)))) | (xor(xor(IN15, !(xor(xor((IN21 | IN6) | (!(IN29)), true), !(IN11 | IN16)))), !(IN21)))))))

*)

FUNCTION_BLOCK F_CollectInput
  VAR_IN_OUT
      Data : ARRAY[1..50] OF BOOL;
  END_VAR
  VAR_INPUT
      TICK  : BOOL := 0;
      IN1   : BOOL := 0;
      IN2   : BOOL := 0;
      IN3   : BOOL := 0;
      IN4   : BOOL := 0;
      IN5   : BOOL := 0;
      RESET : BOOL := FALSE;
  END_VAR
  VAR_OUTPUT
      Finished : BOOL;
  END_VAR
  VAR
      j    : USINT := 1;
      tock : BOOL  := 0;
  END_VAR
  IF NOT RESET AND tock = NOT TICK THEN
      Data[j]   := IN1;
      Data[j+1] := IN2;
      Data[j+2] := IN3;
      Data[j+3] := IN4;
      Data[j+4] := IN5;
      j := j + 5;
      tock := TICK;
  ELSE
      j := 1;
      tock := 0;
  END_IF;
  Finished := (j > 50);
END_FUNCTION_BLOCK

PROGRAM Boiler
  VAR
    Data  : ARRAY[1..50] OF BOOL;
    Ready : BOOL;
    CollectInput : F_CollectInput;
  END_VAR
  VAR
    TICK     AT %IX1.0 : BOOL;
    IN1      AT %IX0.3 : BOOL;
    IN2      AT %IX0.4 : BOOL;
    IN3      AT %IX0.5 : BOOL;
    IN4      AT %IX0.6 : BOOL;
    IN5      AT %IX0.7 : BOOL;
    OutReady AT %QX0.0 : BOOL := FALSE;
    FeedNext AT %QX0.1 : BOOL := FALSE;
    Out      AT %QX0.2 : BOOL;
  END_VAR
  CollectInput(TICK:=TICK, IN1:=IN1, IN2:=IN2, IN3:=IN3, IN4:=IN4, IN5:=IN5);
  Ready := CollectInput.Finished;
  FeedNext := 1;
  IF Ready THEN
    Out := (((((Data[23] AND Data[50]) OR TRUE) XOR (NOT (((((Data[2] AND (((Data[36] XOR (Data[7] OR Data[13])) XOR ((NOT Data[18]) AND (NOT Data[35]))) OR ((((Data[26] AND Data[39]) AND ((Data[30] XOR Data[3]) XOR Data[8])) XOR ((((Data[44] XOR Data[21]) XOR Data[35]) XOR (Data[13] OR Data[29])) XOR ((Data[6] XOR Data[46]) XOR Data[32]))) XOR ((NOT Data[27]) OR (Data[49] OR Data[27]))))) XOR (NOT (Data[28] OR Data[36]))) XOR Data[31]) XOR (((((((((((Data[26] XOR Data[14]) XOR Data[11]) XOR ((Data[42] XOR Data[50]) XOR Data[34])) XOR Data[29]) XOR (NOT Data[42])) XOR Data[17]) XOR Data[33]) XOR (((Data[2] AND (Data[40] AND Data[9])) XOR (Data[26] AND (Data[23] OR Data[38]))) XOR Data[10])) XOR (((Data[23] OR ((Data[49] XOR Data[18]) XOR Data[18])) OR ((((Data[10] XOR Data[38]) XOR Data[17]) XOR (Data[31] AND Data[19])) XOR (Data[50] OR Data[39]))) OR (NOT (((NOT Data[15]) XOR ((Data[10] XOR Data[30]) XOR Data[41])) XOR Data[17])))) XOR Data[41]) AND (NOT ((Data[23] XOR (Data[34] AND (((Data[7] OR Data[19]) XOR (Data[31] AND Data[35])) XOR (NOT Data[42])))) XOR ((NOT (Data[36] AND Data[35])) AND ((NOT Data[6]) AND (Data[9] OR Data[17]))))))) XOR Data[6]))) XOR ((NOT (((((NOT Data[6]) OR ((Data[19] AND Data[9]) OR (Data[47] OR Data[24]))) OR (((NOT Data[43]) OR ((Data[29] XOR Data[49]) XOR Data[49])) OR Data[34])) OR Data[19]) OR (((NOT ((Data[21] XOR (NOT Data[35])) XOR (NOT (NOT Data[7])))) XOR Data[31]) XOR ((FALSE AND ((Data[27] OR Data[44]) OR Data[9])) OR (((Data[16] OR Data[28]) OR (Data[33] OR Data[40])) OR (NOT Data[34])))))) AND ((NOT (Data[38] OR (Data[30] OR (((((Data[31] XOR Data[2]) XOR Data[4]) OR (Data[29] AND Data[7])) XOR (NOT ((Data[7] XOR FALSE) XOR Data[43]))) XOR (((Data[23] XOR Data[28]) XOR Data[27]) AND Data[20]))))) OR (((NOT (((Data[22] XOR ((Data[45] XOR Data[6]) XOR Data[27])) XOR Data[21]) OR (Data[36] AND (Data[47] AND Data[2])))) AND ((((Data[12] OR Data[27]) AND (Data[27] AND Data[26])) AND (Data[6] OR (Data[3] AND Data[10]))) AND (((Data[44] OR Data[37]) OR (Data[17] OR Data[19])) OR (((Data[11] AND Data[29]) XOR Data[2]) XOR (NOT Data[40]))))) AND ((((((Data[50] XOR Data[4]) XOR Data[25]) OR (NOT Data[12])) OR (((Data[13] OR Data[7]) XOR (Data[10] AND Data[39])) XOR Data[47])) OR TRUE) OR (((((((Data[27] OR Data[11]) XOR (Data[42] AND Data[28])) XOR (Data[19] OR Data[24])) XOR FALSE) XOR ((Data[28] OR Data[32]) OR (NOT Data[49]))) XOR (NOT Data[50])) XOR ((NOT ((Data[40] XOR Data[5]) XOR Data[7])) AND (NOT Data[40])))))))) AND ((((NOT ((NOT (((NOT ((Data[34] XOR Data[33]) XOR Data[17])) OR ((Data[20] AND Data[38]) AND (Data[39] AND Data[6]))) AND (Data[12] AND (NOT ((Data[9] XOR Data[5]) XOR Data[8]))))) AND ((((Data[11] XOR (NOT (((Data[50] OR Data[26]) XOR (NOT Data[33])) XOR Data[14]))) XOR Data[32]) XOR (((NOT (Data[27] OR Data[20])) AND (((NOT Data[38]) XOR (Data[14] OR Data[18])) XOR (Data[30] AND Data[44]))) AND (NOT ((Data[45] AND Data[35]) AND (Data[28] AND Data[49]))))) XOR ((Data[8] XOR ((NOT ((Data[48] XOR Data[20]) XOR Data[10])) OR Data[9])) XOR ((NOT (NOT Data[28])) AND (((Data[17] AND Data[28]) XOR (NOT Data[35])) XOR (Data[9] OR Data[18]))))))) XOR (Data[41] OR (NOT ((((NOT ((Data[5] AND Data[1]) OR ((Data[50] XOR Data[32]) XOR Data[38]))) AND TRUE) XOR (((((NOT ((Data[11] XOR Data[43]) XOR Data[38])) XOR ((((Data[49] XOR Data[30]) XOR Data[35]) XOR (Data[34] AND Data[33])) XOR (Data[19] OR Data[27]))) XOR ((Data[9] AND Data[18]) AND ((FALSE XOR Data[7]) XOR Data[40]))) XOR ((((Data[15] OR Data[48]) XOR Data[45]) XOR (NOT Data[47])) OR ((NOT Data[44]) AND (NOT Data[21])))) XOR ((((Data[15] OR Data[44]) AND (NOT Data[2])) XOR ((Data[10] OR Data[4]) OR (NOT Data[14]))) XOR FALSE))) XOR Data[8])))) XOR Data[12]) AND (((((((Data[28] XOR (NOT ((Data[36] XOR (Data[8] AND (Data[6] OR Data[28]))) XOR ((((Data[44] XOR Data[8]) XOR Data[44]) XOR (Data[16] OR Data[15])) XOR (Data[36] OR Data[22]))))) XOR Data[40]) AND ((((Data[8] XOR (((Data[48] OR Data[38]) OR ((Data[40] XOR Data[46]) XOR Data[32])) OR (((Data[15] XOR Data[16]) XOR Data[46]) OR Data[25]))) XOR (NOT (NOT (NOT Data[17])))) XOR (((((Data[1] OR Data[16]) AND (Data[2] OR Data[15])) AND (NOT Data[19])) XOR (((Data[42] OR Data[44]) OR Data[35]) AND (NOT (Data[48] OR Data[35])))) XOR Data[3])) XOR (((((Data[9] AND Data[26]) AND ((Data[1] XOR Data[30]) XOR Data[16])) AND (Data[9] OR ((Data[4] XOR Data[44]) XOR Data[15]))) XOR ((NOT ((Data[47] XOR Data[5]) XOR Data[41])) AND (Data[18] OR ((Data[9] XOR Data[45]) XOR Data[23])))) XOR (NOT Data[32])))) XOR (((((NOT Data[27]) XOR Data[9]) XOR (((Data[16] XOR (Data[41] OR Data[36])) XOR Data[41]) OR ((Data[48] XOR Data[22]) XOR (Data[25] AND Data[36])))) OR (NOT (Data[46] AND (((Data[16] XOR Data[48]) XOR Data[39]) OR ((Data[15] XOR TRUE) XOR Data[12]))))) OR Data[44])) XOR (Data[48] AND ((NOT (NOT ((Data[27] AND Data[33]) AND (Data[33] AND Data[39])))) OR (Data[19] AND Data[41])))) XOR (NOT Data[40])) XOR (NOT ((((((((((Data[30] OR Data[38]) XOR ((Data[39] XOR Data[19]) XOR Data[33])) XOR (Data[40] OR Data[13])) XOR Data[44]) XOR ((NOT Data[26]) AND Data[23])) XOR (((Data[16] OR Data[48]) AND Data[22]) OR (Data[23] AND (Data[1] AND Data[3])))) XOR Data[8]) XOR ((NOT ((Data[43] AND Data[11]) AND Data[33])) AND Data[16])) XOR ((NOT (((Data[47] XOR Data[34]) XOR Data[37]) OR (NOT Data[19]))) OR ((NOT Data[27]) AND (((Data[3] XOR Data[37]) XOR Data[48]) OR Data[22])))) OR ((Data[15] XOR (NOT ((((Data[21] OR Data[6]) OR (NOT Data[29])) XOR TRUE) XOR (NOT (Data[11] OR Data[16]))))) XOR (NOT Data[21])))))));
    OutReady := 1;
    CollectInput(RESET:=TRUE);
  END_IF;
END_PROGRAM

CONFIGURATION Config0
  RESOURCE Res0 ON PLC
    TASK task0(INTERVAL := T#20ms,PRIORITY := 0);
    PROGRAM instance0 WITH task0 : Boiler;
  END_RESOURCE
END_CONFIGURATION

(* ---- RND-EXPR_rebox-pedal-toons.st ---- *)
(*
This code implements a randomly grown symbolic expression:

IN6 & IN4

*)

FUNCTION_BLOCK F_CollectInput
  VAR_IN_OUT
      Data : ARRAY[1..50] OF BOOL;
  END_VAR
  VAR_INPUT
      TICK  : BOOL := 0;
      IN1   : BOOL := 0;
      IN2   : BOOL := 0;
      IN3   : BOOL := 0;
      IN4   : BOOL := 0;
      IN5   : BOOL := 0;
      RESET : BOOL := FALSE;
  END_VAR
  VAR_OUTPUT
      Finished : BOOL;
  END_VAR
  VAR
      j    : USINT := 1;
      tock : BOOL  := 0;
  END_VAR
  IF NOT RESET AND tock = NOT TICK THEN
      Data[j]   := IN1;
      Data[j+1] := IN2;
      Data[j+2] := IN3;
      Data[j+3] := IN4;
      Data[j+4] := IN5;
      j := j + 5;
      tock := TICK;
  ELSE
      j := 1;
      tock := 0;
  END_IF;
  Finished := (j > 50);
END_FUNCTION_BLOCK

PROGRAM Boiler
  VAR
    Data  : ARRAY[1..50] OF BOOL;
    Ready : BOOL;
    CollectInput : F_CollectInput;
  END_VAR
  VAR
    TICK     AT %IX1.0 : BOOL;
    IN1      AT %IX0.3 : BOOL;
    IN2      AT %IX0.4 : BOOL;
    IN3      AT %IX0.5 : BOOL;
    IN4      AT %IX0.6 : BOOL;
    IN5      AT %IX0.7 : BOOL;
    OutReady AT %QX0.0 : BOOL := FALSE;
    FeedNext AT %QX0.1 : BOOL := FALSE;
    Out      AT %QX0.2 : BOOL;
  END_VAR
  CollectInput(TICK:=TICK, IN1:=IN1, IN2:=IN2, IN3:=IN3, IN4:=IN4, IN5:=IN5);
  Ready := CollectInput.Finished;
  FeedNext := 1;
  IF Ready THEN
    Out := (Data[6] AND Data[4]);
    OutReady := 1;
    CollectInput(RESET:=TRUE);
  END_IF;
END_PROGRAM

CONFIGURATION Config0
  RESOURCE Res0 ON PLC
    TASK task0(INTERVAL := T#20ms,PRIORITY := 0);
    PROGRAM instance0 WITH task0 : Boiler;
  END_RESOURCE
END_CONFIGURATION

(* ---- RND-EXPR_regal-dowry-slake.st ---- *)
(*
This code implements a randomly grown symbolic expression:

((((xor(xor((!(!(xor(xor(IN29 | IN28, IN36), IN43 | IN8)))) & ((((xor(xor(IN27, IN14), IN33)) & (xor(xor(IN48, IN39), IN30))) | (IN41 | (xor(xor(false, IN35), IN14)))) & ((xor(xor(IN31, IN4 & IN24), IN26)) & (xor(xor(IN3 & IN41, !(IN32)), IN4 & IN8)))), !(IN48)), ((!(!(IN1 & IN47))) | IN45) | (IN26 & ((true | (xor(xor(IN20, IN1), IN45))) | ((xor(xor(false, IN37), IN14)) | (IN19 & IN30)))))) | IN41) | (xor(xor((IN9 | (xor(xor(!((xor(xor(IN13, false), IN29)) & (IN18 | IN23)), (xor(xor(IN33 | IN25, !(IN41)), xor(xor(IN43, IN27), IN33))) & ((true | IN30) | (IN19 | IN42))), true & (xor(xor(IN38 | IN12, xor(xor(IN10, false), IN5)), IN16 & IN45))))) & IN40, IN44), !(!(!((!(IN8 | IN20)) & IN38)))))) & (xor(xor((!(!(!(!((IN37 & IN4) & (xor(xor(IN34, false), false))))))) | (((!(!((IN48 | IN10) & (IN45 & IN23)))) & ((!(!(!(IN49)))) | true)) & (xor(xor((xor(xor((!(IN33)) | (IN25 | IN11), IN7), IN37)) & ((!(IN24 & IN11)) | (xor(xor(IN27 | IN38, IN13), false))), xor(xor(IN36, IN31), (xor(xor(true, IN42), !(IN15))) | ((IN6 | IN45) | (IN36 | IN4)))), IN11))), !(!(((xor(xor(IN20 | (!(IN38)), xor(xor(IN50 | IN24, IN46 | IN36), !(IN40))), (IN49 | IN28) & (xor(xor(IN1, IN12), IN31)))) | (!(IN18))) & (!(IN21 & ((xor(xor(IN1, IN6), IN21)) & (!(IN41)))))))), true))) & (!((((IN7 | (xor(xor(((xor(xor(IN10, IN19), IN23)) & (xor(xor(IN1, IN21), IN36))) & (!(xor(xor(IN44, IN49), IN18))), IN32), IN47))) & (((IN4 & (!(IN44))) | false) & (!(IN47)))) & (xor(xor(xor(xor(((xor(xor(IN46, IN15 | IN27), IN46 & IN21)) | (xor(xor(xor(xor(IN31, IN24), IN28), xor(xor(IN1, IN25), IN11)), xor(xor(IN4, true), IN19)))) & IN27, IN46), !(((IN19 & IN18) & (!(IN14))) | ((xor(xor(IN2, IN6), IN21)) & IN40))), (xor(xor(xor(xor(xor(xor(!(IN12), IN39 | IN10), !(IN37)), xor(xor(xor(xor(true, IN48), IN48), xor(xor(IN2, IN29), IN49)), IN25 | IN31)), xor(xor(IN42 & IN17, IN30 | IN2), IN43)), xor(xor((IN43 | IN20) | (IN35 | IN17), (!(IN43)) & (xor(xor(IN3, IN36), IN10))), !(IN47 & IN47))), xor(xor(xor(xor(IN11 | IN13, !(IN43)), xor(xor(IN39, IN17), IN39)), xor(xor(xor(xor(IN42, IN45), IN22), !(IN24)), xor(xor(IN29, IN18), IN50))), !(IN43 & IN18)))) & (((!(!(IN42))) & (xor(xor(false, IN15 | IN35), xor(xor(IN5, IN14), IN47)))) & (!(IN32)))), ((xor(xor((xor(xor(IN13, IN12), IN19)) & (IN35 | IN49), xor(xor(xor(xor(IN15, IN39), IN44), IN36), IN12)), xor(xor(!(IN34), IN4 | true), xor(xor(IN30, IN43), IN22)))) & IN18) | ((!((IN26 & IN23) & IN34)) | ((xor(xor(IN3 | IN31, xor(xor(IN34, IN44), IN20)), xor(xor(IN15, IN38), IN47))) & (!(IN22))))))) & (xor(xor((!((xor(xor(xor(xor(!(IN14), !(IN12)), !(IN33)), xor(xor(IN3, xor(xor(IN43, IN21), IN10)), xor(xor(IN38, IN46), IN29))), IN39)) & (((xor(xor(IN17, IN6), IN11)) | (xor(xor(IN32, IN41), IN31))) & (xor(xor(IN39 & IN5, true), !(IN5)))))) | (!(IN33)), xor(xor(IN49 | ((((IN25 & IN33) | (IN12 & IN39)) | ((xor(xor(IN30, IN11), IN41)) | IN22)) | (((!(IN36)) & (false & IN25)) | (xor(xor(IN18 | IN14, IN36), IN7 | IN49)))), !(IN50)), ((!(!(IN28))) & (!(!(IN49 & IN47)))) & IN50)), IN21))))

*)

FUNCTION_BLOCK F_CollectInput
  VAR_IN_OUT
      Data : ARRAY[1..50] OF BOOL;
  END_VAR
  VAR_INPUT
      TICK  : BOOL := 0;
      IN1   : BOOL := 0;
      IN2   : BOOL := 0;
      IN3   : BOOL := 0;
      IN4   : BOOL := 0;
      IN5   : BOOL := 0;
      RESET : BOOL := FALSE;
  END_VAR
  VAR_OUTPUT
      Finished : BOOL;
  END_VAR
  VAR
      j    : USINT := 1;
      tock : BOOL  := 0;
  END_VAR
  IF NOT RESET AND tock = NOT TICK THEN
      Data[j]   := IN1;
      Data[j+1] := IN2;
      Data[j+2] := IN3;
      Data[j+3] := IN4;
      Data[j+4] := IN5;
      j := j + 5;
      tock := TICK;
  ELSE
      j := 1;
      tock := 0;
  END_IF;
  Finished := (j > 50);
END_FUNCTION_BLOCK

PROGRAM Boiler
  VAR
    Data  : ARRAY[1..50] OF BOOL;
    Ready : BOOL;
    CollectInput : F_CollectInput;
  END_VAR
  VAR
    TICK     AT %IX1.0 : BOOL;
    IN1      AT %IX0.3 : BOOL;
    IN2      AT %IX0.4 : BOOL;
    IN3      AT %IX0.5 : BOOL;
    IN4      AT %IX0.6 : BOOL;
    IN5      AT %IX0.7 : BOOL;
    OutReady AT %QX0.0 : BOOL := FALSE;
    FeedNext AT %QX0.1 : BOOL := FALSE;
    Out      AT %QX0.2 : BOOL;
  END_VAR
  CollectInput(TICK:=TICK, IN1:=IN1, IN2:=IN2, IN3:=IN3, IN4:=IN4, IN5:=IN5);
  Ready := CollectInput.Finished;
  FeedNext := 1;
  IF Ready THEN
    Out := ((((((((NOT (NOT (((Data[29] OR Data[28]) XOR Data[36]) XOR (Data[43] OR Data[8])))) AND (((((Data[27] XOR Data[14]) XOR Data[33]) AND ((Data[48] XOR Data[39]) XOR Data[30])) OR (Data[41] OR ((FALSE XOR Data[35]) XOR Data[14]))) AND (((Data[31] XOR (Data[4] AND Data[24])) XOR Data[26]) AND (((Data[3] AND Data[41]) XOR (NOT Data[32])) XOR (Data[4] AND Data[8]))))) XOR (NOT Data[48])) XOR (((NOT (NOT (Data[1] AND Data[47]))) OR Data[45]) OR (Data[26] AND ((TRUE OR ((Data[20] XOR Data[1]) XOR Data[45])) OR (((FALSE XOR Data[37]) XOR Data[14]) OR (Data[19] AND Data[30])))))) OR Data[41]) OR ((((Data[9] OR (((NOT (((Data[13] XOR FALSE) XOR Data[29]) AND (Data[18] OR Data[23]))) XOR ((((Data[33] OR Data[25]) XOR (NOT Data[41])) XOR ((Data[43] XOR Data[27]) XOR Data[33])) AND ((TRUE OR Data[30]) OR (Data[19] OR Data[42])))) XOR (TRUE AND (((Data[38] OR Data[12]) XOR ((Data[10] XOR FALSE) XOR Data[5])) XOR (Data[16] AND Data[45]))))) AND Data[40]) XOR Data[44]) XOR (NOT (NOT (NOT ((NOT (Data[8] OR Data[20])) AND Data[38])))))) AND ((((NOT (NOT (NOT (NOT ((Data[37] AND Data[4]) AND ((Data[34] XOR FALSE) XOR FALSE)))))) OR (((NOT (NOT ((Data[48] OR Data[10]) AND (Data[45] AND Data[23])))) AND ((NOT (NOT (NOT Data[49]))) OR TRUE)) AND (((((((NOT Data[33]) OR (Data[25] OR Data[11])) XOR Data[7]) XOR Data[37]) AND ((NOT (Data[24] AND Data[11])) OR (((Data[27] OR Data[38]) XOR Data[13]) XOR FALSE))) XOR ((Data[36] XOR Data[31]) XOR (((TRUE XOR Data[42]) XOR (NOT Data[15])) OR ((Data[6] OR Data[45]) OR (Data[36] OR Data[4]))))) XOR Data[11]))) XOR (NOT (NOT (((((Data[20] OR (NOT Data[38])) XOR (((Data[50] OR Data[24]) XOR (Data[46] OR Data[36])) XOR (NOT Data[40]))) XOR ((Data[49] OR Data[28]) AND ((Data[1] XOR Data[12]) XOR Data[31]))) OR (NOT Data[18])) AND (NOT (Data[21] AND (((Data[1] XOR Data[6]) XOR Data[21]) AND (NOT Data[41])))))))) XOR TRUE)) AND (NOT ((((Data[7] OR ((((((Data[10] XOR Data[19]) XOR Data[23]) AND ((Data[1] XOR Data[21]) XOR Data[36])) AND (NOT ((Data[44] XOR Data[49]) XOR Data[18]))) XOR Data[32]) XOR Data[47])) AND (((Data[4] AND (NOT Data[44])) OR FALSE) AND (NOT Data[47]))) AND ((((((((Data[46] XOR (Data[15] OR Data[27])) XOR (Data[46] AND Data[21])) OR ((((Data[31] XOR Data[24]) XOR Data[28]) XOR ((Data[1] XOR Data[25]) XOR Data[11])) XOR ((Data[4] XOR TRUE) XOR Data[19]))) AND Data[27]) XOR Data[46]) XOR (NOT (((Data[19] AND Data[18]) AND (NOT Data[14])) OR (((Data[2] XOR Data[6]) XOR Data[21]) AND Data[40])))) XOR ((((((((NOT Data[12]) XOR (Data[39] OR Data[10])) XOR (NOT Data[37])) XOR ((((TRUE XOR Data[48]) XOR Data[48]) XOR ((Data[2] XOR Data[29]) XOR Data[49])) XOR (Data[25] OR Data[31]))) XOR (((Data[42] AND Data[17]) XOR (Data[30] OR Data[2])) XOR Data[43])) XOR ((((Data[43] OR Data[20]) OR (Data[35] OR Data[17])) XOR ((NOT Data[43]) AND ((Data[3] XOR Data[36]) XOR Data[10]))) XOR (NOT (Data[47] AND Data[47])))) XOR (((((Data[11] OR Data[13]) XOR (NOT Data[43])) XOR ((Data[39] XOR Data[17]) XOR Data[39])) XOR ((((Data[42] XOR Data[45]) XOR Data[22]) XOR (NOT Data[24])) XOR ((Data[29] XOR Data[18]) XOR Data[50]))) XOR (NOT (Data[43] AND Data[18])))) AND (((NOT (NOT Data[42])) AND ((FALSE XOR (Data[15] OR Data[35])) XOR ((Data[5] XOR Data[14]) XOR Data[47]))) AND (NOT Data[32])))) XOR (((((((Data[13] XOR Data[12]) XOR Data[19]) AND (Data[35] OR Data[49])) XOR ((((Data[15] XOR Data[39]) XOR Data[44]) XOR Data[36]) XOR Data[12])) XOR (((NOT Data[34]) XOR (Data[4] OR TRUE)) XOR ((Data[30] XOR Data[43]) XOR Data[22]))) AND Data[18]) OR ((NOT ((Data[26] AND Data[23]) AND Data[34])) OR ((((Data[3] OR Data[31]) XOR ((Data[34] XOR Data[44]) XOR Data[20])) XOR ((Data[15] XOR Data[38]) XOR Data[47])) AND (NOT Data[22])))))) AND ((((NOT ((((((NOT Data[14]) XOR (NOT Data[12])) XOR (NOT Data[33])) XOR ((Data[3] XOR ((Data[43] XOR Data[21]) XOR Data[10])) XOR ((Data[38] XOR Data[46]) XOR Data[29]))) XOR Data[39]) AND ((((Data[17] XOR Data[6]) XOR Data[11]) OR ((Data[32] XOR Data[41]) XOR Data[31])) AND (((Data[39] AND Data[5]) XOR TRUE) XOR (NOT Data[5]))))) OR (NOT Data[33])) XOR (((Data[49] OR ((((Data[25] AND Data[33]) OR (Data[12] AND Data[39])) OR (((Data[30] XOR Data[11]) XOR Data[41]) OR Data[22])) OR (((NOT Data[36]) AND (FALSE AND Data[25])) OR (((Data[18] OR Data[14]) XOR Data[36]) XOR (Data[7] OR Data[49]))))) XOR (NOT Data[50])) XOR (((NOT (NOT Data[28])) AND (NOT (NOT (Data[49] AND Data[47])))) AND Data[50]))) XOR Data[21]))));
    OutReady := 1;
    CollectInput(RESET:=TRUE);
  END_IF;
END_PROGRAM

CONFIGURATION Config0
  RESOURCE Res0 ON PLC
    TASK task0(INTERVAL := T#20ms,PRIORITY := 0);
    PROGRAM instance0 WITH task0 : Boiler;
  END_RESOURCE
END_CONFIGURATION

(* ---- RND-EXPR_renew-pivot-middy.st ---- *)
(*
This code implements a randomly grown symbolic expression:

IN23 | ((xor(xor(((!((!(!(xor(xor(IN3, IN39), IN23)))) & (xor(xor((IN37 & IN30) | IN33, IN16 | (IN49 | IN9)), xor(xor(IN13 | IN6, !(IN46)), !(IN11)))))) | (!(!(((xor(xor(IN20, IN44), IN17)) & IN43) | (true & IN41))))) | ((!(IN3)) | (!(IN43))), IN3), IN29 & ((xor(xor(xor(xor(IN47, xor(xor((IN37 & IN14) & (!(IN4)), IN41), (IN33 | IN20) | (!(IN39)))), (!(!(IN2))) & (xor(xor(IN38, xor(xor(IN22, IN35), IN46)), IN40))), (!(IN48)) | (xor(xor(IN26 | (true & IN3), !(IN27 & IN36)), IN46))), (IN43 & IN46) | (IN45 | (IN1 | (IN35 | IN6))))) & (xor(xor(!(IN30 | (xor(xor(IN6 | IN23, xor(xor(IN5, IN13), IN16)), IN28 & IN47))), xor(xor((xor(xor(!(IN7), IN8 & IN25), !(IN37))) & (xor(xor(IN3 | IN16, xor(xor(IN15, IN12), IN36)), IN31 | IN30)), IN45 & (xor(xor(IN23 & IN2, IN19 & IN20), IN29))), xor(xor(xor(xor(IN30, !(IN36)), IN6 | IN24), !(IN23 & IN40)), !(IN21)))), xor(xor(!(IN21 | (IN47 | IN1)), ((!(IN40)) & (!(IN48))) & (!(IN16 & IN43))), xor(xor((xor(xor(IN3, IN26), IN3)) | (IN48 | IN43), !(IN41 & IN41)), !(IN38 | IN9)))))))) | (xor(xor(!(!((xor(xor((xor(xor(IN22 & IN18, IN40 & IN17), xor(xor(IN4, IN35), IN12))) | ((IN7 & IN12) | (!(IN34))), ((!(IN3)) | (IN30 | true)) & (!(!(IN33)))), ((IN25 | IN5) & (xor(xor(IN8, IN3), IN47))) & (xor(xor(IN42 | IN9, IN1 | IN39), IN47 | IN50)))) | (!(IN46)))), IN41 | ((!(!(IN12))) & (xor(xor(!((!(!(IN39))) | (xor(xor(xor(xor(IN26, IN22), IN46), xor(xor(IN12, IN37), IN36)), !(IN5)))), ((false & (IN42 | false)) | (!(!(IN14)))) | (xor(xor((IN26 | IN15) & (IN18 | IN11), !(xor(xor(IN49, IN9), IN43))), xor(xor(IN1 & IN37, xor(xor(IN17, IN14), true)), xor(xor(IN25, IN9), IN12))))), !(xor(xor((!(IN15)) | (!(IN2)), IN36), !(IN45 | IN43))))))), (!((((!(xor(xor(IN10, IN25), IN1))) | IN35) | (xor(xor((!(IN20)) & IN36, (IN18 & IN18) & (IN18 & IN20)), IN4 | false))) & ((xor(xor(xor(xor(xor(xor(IN49, IN15), IN11), IN45 & IN14), IN50 & IN46), (true & IN9) | (xor(xor(IN32, IN36), IN25))), (xor(xor(IN28, IN34), IN46)) | (IN49 | IN18))) & ((xor(xor(xor(xor(IN19, IN37), IN17), IN2), IN26 & IN16)) & ((!(IN32)) & IN19))))) & (!(IN35)))))

*)

FUNCTION_BLOCK F_CollectInput
  VAR_IN_OUT
      Data : ARRAY[1..50] OF BOOL;
  END_VAR
  VAR_INPUT
      TICK  : BOOL := 0;
      IN1   : BOOL := 0;
      IN2   : BOOL := 0;
      IN3   : BOOL := 0;
      IN4   : BOOL := 0;
      IN5   : BOOL := 0;
      RESET : BOOL := FALSE;
  END_VAR
  VAR_OUTPUT
      Finished : BOOL;
  END_VAR
  VAR
      j    : USINT := 1;
      tock : BOOL  := 0;
  END_VAR
  IF NOT RESET AND tock = NOT TICK THEN
      Data[j]   := IN1;
      Data[j+1] := IN2;
      Data[j+2] := IN3;
      Data[j+3] := IN4;
      Data[j+4] := IN5;
      j := j + 5;
      tock := TICK;
  ELSE
      j := 1;
      tock := 0;
  END_IF;
  Finished := (j > 50);
END_FUNCTION_BLOCK

PROGRAM Boiler
  VAR
    Data  : ARRAY[1..50] OF BOOL;
    Ready : BOOL;
    CollectInput : F_CollectInput;
  END_VAR
  VAR
    TICK     AT %IX1.0 : BOOL;
    IN1      AT %IX0.3 : BOOL;
    IN2      AT %IX0.4 : BOOL;
    IN3      AT %IX0.5 : BOOL;
    IN4      AT %IX0.6 : BOOL;
    IN5      AT %IX0.7 : BOOL;
    OutReady AT %QX0.0 : BOOL := FALSE;
    FeedNext AT %QX0.1 : BOOL := FALSE;
    Out      AT %QX0.2 : BOOL;
  END_VAR
  CollectInput(TICK:=TICK, IN1:=IN1, IN2:=IN2, IN3:=IN3, IN4:=IN4, IN5:=IN5);
  Ready := CollectInput.Finished;
  FeedNext := 1;
  IF Ready THEN
    Out := (Data[23] OR ((((((NOT ((NOT (NOT ((Data[3] XOR Data[39]) XOR Data[23]))) AND ((((Data[37] AND Data[30]) OR Data[33]) XOR (Data[16] OR (Data[49] OR Data[9]))) XOR (((Data[13] OR Data[6]) XOR (NOT Data[46])) XOR (NOT Data[11]))))) OR (NOT (NOT ((((Data[20] XOR Data[44]) XOR Data[17]) AND Data[43]) OR (TRUE AND Data[41]))))) OR ((NOT Data[3]) OR (NOT Data[43]))) XOR Data[3]) XOR (Data[29] AND (((((Data[47] XOR ((((Data[37] AND Data[14]) AND (NOT Data[4])) XOR Data[41]) XOR ((Data[33] OR Data[20]) OR (NOT Data[39])))) XOR ((NOT (NOT Data[2])) AND ((Data[38] XOR ((Data[22] XOR Data[35]) XOR Data[46])) XOR Data[40]))) XOR ((NOT Data[48]) OR (((Data[26] OR (TRUE AND Data[3])) XOR (NOT (Data[27] AND Data[36]))) XOR Data[46]))) XOR ((Data[43] AND Data[46]) OR (Data[45] OR (Data[1] OR (Data[35] OR Data[6]))))) AND (((NOT (Data[30] OR (((Data[6] OR Data[23]) XOR ((Data[5] XOR Data[13]) XOR Data[16])) XOR (Data[28] AND Data[47])))) XOR ((((((NOT Data[7]) XOR (Data[8] AND Data[25])) XOR (NOT Data[37])) AND (((Data[3] OR Data[16]) XOR ((Data[15] XOR Data[12]) XOR Data[36])) XOR (Data[31] OR Data[30]))) XOR (Data[45] AND (((Data[23] AND Data[2]) XOR (Data[19] AND Data[20])) XOR Data[29]))) XOR ((((Data[30] XOR (NOT Data[36])) XOR (Data[6] OR Data[24])) XOR (NOT (Data[23] AND Data[40]))) XOR (NOT Data[21])))) XOR (((NOT (Data[21] OR (Data[47] OR Data[1]))) XOR (((NOT Data[40]) AND (NOT Data[48])) AND (NOT (Data[16] AND Data[43])))) XOR (((((Data[3] XOR Data[26]) XOR Data[3]) OR (Data[48] OR Data[43])) XOR (NOT (Data[41] AND Data[41]))) XOR (NOT (Data[38] OR Data[9])))))))) OR (((NOT (NOT (((((((Data[22] AND Data[18]) XOR (Data[40] AND Data[17])) XOR ((Data[4] XOR Data[35]) XOR Data[12])) OR ((Data[7] AND Data[12]) OR (NOT Data[34]))) XOR (((NOT Data[3]) OR (Data[30] OR TRUE)) AND (NOT (NOT Data[33])))) XOR (((Data[25] OR Data[5]) AND ((Data[8] XOR Data[3]) XOR Data[47])) AND (((Data[42] OR Data[9]) XOR (Data[1] OR Data[39])) XOR (Data[47] OR Data[50])))) OR (NOT Data[46])))) XOR (Data[41] OR ((NOT (NOT Data[12])) AND (((NOT ((NOT (NOT Data[39])) OR ((((Data[26] XOR Data[22]) XOR Data[46]) XOR ((Data[12] XOR Data[37]) XOR Data[36])) XOR (NOT Data[5])))) XOR (((FALSE AND (Data[42] OR FALSE)) OR (NOT (NOT Data[14]))) OR ((((Data[26] OR Data[15]) AND (Data[18] OR Data[11])) XOR (NOT ((Data[49] XOR Data[9]) XOR Data[43]))) XOR (((Data[1] AND Data[37]) XOR ((Data[17] XOR Data[14]) XOR TRUE)) XOR ((Data[25] XOR Data[9]) XOR Data[12]))))) XOR (NOT ((((NOT Data[15]) OR (NOT Data[2])) XOR Data[36]) XOR (NOT (Data[45] OR Data[43])))))))) XOR ((NOT ((((NOT ((Data[10] XOR Data[25]) XOR Data[1])) OR Data[35]) OR ((((NOT Data[20]) AND Data[36]) XOR ((Data[18] AND Data[18]) AND (Data[18] AND Data[20]))) XOR (Data[4] OR FALSE))) AND (((((((Data[49] XOR Data[15]) XOR Data[11]) XOR (Data[45] AND Data[14])) XOR (Data[50] AND Data[46])) XOR ((TRUE AND Data[9]) OR ((Data[32] XOR Data[36]) XOR Data[25]))) XOR (((Data[28] XOR Data[34]) XOR Data[46]) OR (Data[49] OR Data[18]))) AND (((((Data[19] XOR Data[37]) XOR Data[17]) XOR Data[2]) XOR (Data[26] AND Data[16])) AND ((NOT Data[32]) AND Data[19]))))) AND (NOT Data[35])))));
    OutReady := 1;
    CollectInput(RESET:=TRUE);
  END_IF;
END_PROGRAM

CONFIGURATION Config0
  RESOURCE Res0 ON PLC
    TASK task0(INTERVAL := T#20ms,PRIORITY := 0);
    PROGRAM instance0 WITH task0 : Boiler;
  END_RESOURCE
END_CONFIGURATION

(* ---- RND-EXPR_rives-flume-hires.st ---- *)
(*
This code implements a randomly grown symbolic expression:

!(!(xor(xor(!((IN33 | ((xor(xor(!(xor(xor(IN35, IN28), IN41)), xor(xor(xor(xor(IN11, IN2), IN21), IN44), xor(xor(IN22, IN2), IN29))), !(IN43))) & ((IN14 | (xor(xor(IN4, false), IN29))) | ((xor(xor(IN40, IN17), IN18)) & IN4)))) & (IN1 & (((xor(xor(xor(xor(IN44, IN36), IN38), IN7 & IN41), IN26 & IN16)) | ((!(IN35)) | (!(IN26)))) & IN50))), IN37 | IN14), IN39)))

*)

FUNCTION_BLOCK F_CollectInput
  VAR_IN_OUT
      Data : ARRAY[1..50] OF BOOL;
  END_VAR
  VAR_INPUT
      TICK  : BOOL := 0;
      IN1   : BOOL := 0;
      IN2   : BOOL := 0;
      IN3   : BOOL := 0;
      IN4   : BOOL := 0;
      IN5   : BOOL := 0;
      RESET : BOOL := FALSE;
  END_VAR
  VAR_OUTPUT
      Finished : BOOL;
  END_VAR
  VAR
      j    : USINT := 1;
      tock : BOOL  := 0;
  END_VAR
  IF NOT RESET AND tock = NOT TICK THEN
      Data[j]   := IN1;
      Data[j+1] := IN2;
      Data[j+2] := IN3;
      Data[j+3] := IN4;
      Data[j+4] := IN5;
      j := j + 5;
      tock := TICK;
  ELSE
      j := 1;
      tock := 0;
  END_IF;
  Finished := (j > 50);
END_FUNCTION_BLOCK

PROGRAM Boiler
  VAR
    Data  : ARRAY[1..50] OF BOOL;
    Ready : BOOL;
    CollectInput : F_CollectInput;
  END_VAR
  VAR
    TICK     AT %IX1.0 : BOOL;
    IN1      AT %IX0.3 : BOOL;
    IN2      AT %IX0.4 : BOOL;
    IN3      AT %IX0.5 : BOOL;
    IN4      AT %IX0.6 : BOOL;
    IN5      AT %IX0.7 : BOOL;
    OutReady AT %QX0.0 : BOOL := FALSE;
    FeedNext AT %QX0.1 : BOOL := FALSE;
    Out      AT %QX0.2 : BOOL;
  END_VAR
  CollectInput(TICK:=TICK, IN1:=IN1, IN2:=IN2, IN3:=IN3, IN4:=IN4, IN5:=IN5);
  Ready := CollectInput.Finished;
  FeedNext := 1;
  IF Ready THEN
    Out := (NOT (NOT (((NOT ((Data[33] OR ((((NOT ((Data[35] XOR Data[28]) XOR Data[41])) XOR ((((Data[11] XOR Data[2]) XOR Data[21]) XOR Data[44]) XOR ((Data[22] XOR Data[2]) XOR Data[29]))) XOR (NOT Data[43])) AND ((Data[14] OR ((Data[4] XOR FALSE) XOR Data[29])) OR (((Data[40] XOR Data[17]) XOR Data[18]) AND Data[4])))) AND (Data[1] AND ((((((Data[44] XOR Data[36]) XOR Data[38]) XOR (Data[7] AND Data[41])) XOR (Data[26] AND Data[16])) OR ((NOT Data[35]) OR (NOT Data[26]))) AND Data[50])))) XOR (Data[37] OR Data[14])) XOR Data[39])));
    OutReady := 1;
    CollectInput(RESET:=TRUE);
  END_IF;
END_PROGRAM

CONFIGURATION Config0
  RESOURCE Res0 ON PLC
    TASK task0(INTERVAL := T#20ms,PRIORITY := 0);
    PROGRAM instance0 WITH task0 : Boiler;
  END_RESOURCE
END_CONFIGURATION
